(* IEC 61131-3 sources: STAR-PLC-Agent/results/raw/four_group_20261114/star_terra/PUB008/generation/sim_00, 1 file *)

(* ---- test_program.st ---- *)
PROGRAM PLC_PRG
VAR
 BenchStep : UDINT := 0;
 BenchCalls : UDINT := 0;
 BenchDone : BOOL := FALSE;
 BenchUut0 : FB_Task;
 BenchUut1 : FB_Task;
 Binding_0_analogValues : ARRAY[1..14] OF INT;
 Binding_0_channels : ARRAY[1..14] OF ST_AnalogChannel;
 Binding_1_analogValues : ARRAY[1..10] OF INT;
 Binding_1_channels : ARRAY[1..9] OF ST_AnalogChannel;
 TraceIn_count : ARRAY[0..3] OF DINT;
 TraceOut_analogValues_1 : ARRAY[0..3] OF INT;
 TraceOut_analogValues_2 : ARRAY[0..3] OF INT;
 TraceOut_analogValues_3 : ARRAY[0..3] OF INT;
 TraceOut_analogValues_4 : ARRAY[0..3] OF INT;
 TraceOut_analogValues_5 : ARRAY[0..3] OF INT;
 TraceOut_analogValues_6 : ARRAY[0..3] OF INT;
 TraceOut_analogValues_7 : ARRAY[0..3] OF INT;
 TraceOut_analogValues_8 : ARRAY[0..3] OF INT;
 TraceOut_analogValues_9 : ARRAY[0..3] OF INT;
 TraceOut_analogValues_10 : ARRAY[0..3] OF INT;
 TraceOut_analogValues_11 : ARRAY[0..3] OF INT;
 TraceOut_analogValues_12 : ARRAY[0..3] OF INT;
 TraceOut_analogValues_13 : ARRAY[0..3] OF INT;
 TraceOut_analogValues_14 : ARRAY[0..3] OF INT;
 TraceOut_channels_1_enable : ARRAY[0..3] OF BOOL;
 TraceOut_channels_1_hiLIM : ARRAY[0..3] OF REAL;
 TraceOut_channels_1_loLIM : ARRAY[0..3] OF REAL;
 TraceOut_channels_1_bipolar : ARRAY[0..3] OF BOOL;
 TraceOut_channels_1_measuringMode : ARRAY[0..3] OF INT;
 TraceOut_channels_1_retVal : ARRAY[0..3] OF WORD;
 TraceOut_channels_1_outputValue : ARRAY[0..3] OF REAL;
 TraceOut_channels_2_enable : ARRAY[0..3] OF BOOL;
 TraceOut_channels_2_hiLIM : ARRAY[0..3] OF REAL;
 TraceOut_channels_2_loLIM : ARRAY[0..3] OF REAL;
 TraceOut_channels_2_bipolar : ARRAY[0..3] OF BOOL;
 TraceOut_channels_2_measuringMode : ARRAY[0..3] OF INT;
 TraceOut_channels_2_retVal : ARRAY[0..3] OF WORD;
 TraceOut_channels_2_outputValue : ARRAY[0..3] OF REAL;
 TraceOut_channels_3_enable : ARRAY[0..3] OF BOOL;
 TraceOut_channels_3_hiLIM : ARRAY[0..3] OF REAL;
 TraceOut_channels_3_loLIM : ARRAY[0..3] OF REAL;
 TraceOut_channels_3_bipolar : ARRAY[0..3] OF BOOL;
 TraceOut_channels_3_measuringMode : ARRAY[0..3] OF INT;
 TraceOut_channels_3_retVal : ARRAY[0..3] OF WORD;
 TraceOut_channels_3_outputValue : ARRAY[0..3] OF REAL;
 TraceOut_channels_4_enable : ARRAY[0..3] OF BOOL;
 TraceOut_channels_4_hiLIM : ARRAY[0..3] OF REAL;
 TraceOut_channels_4_loLIM : ARRAY[0..3] OF REAL;
 TraceOut_channels_4_bipolar : ARRAY[0..3] OF BOOL;
 TraceOut_channels_4_measuringMode : ARRAY[0..3] OF INT;
 TraceOut_channels_4_retVal : ARRAY[0..3] OF WORD;
 TraceOut_channels_4_outputValue : ARRAY[0..3] OF REAL;
 TraceOut_channels_5_enable : ARRAY[0..3] OF BOOL;
 TraceOut_channels_5_hiLIM : ARRAY[0..3] OF REAL;
 TraceOut_channels_5_loLIM : ARRAY[0..3] OF REAL;
 TraceOut_channels_5_bipolar : ARRAY[0..3] OF BOOL;
 TraceOut_channels_5_measuringMode : ARRAY[0..3] OF INT;
 TraceOut_channels_5_retVal : ARRAY[0..3] OF WORD;
 TraceOut_channels_5_outputValue : ARRAY[0..3] OF REAL;
 TraceOut_channels_6_enable : ARRAY[0..3] OF BOOL;
 TraceOut_channels_6_hiLIM : ARRAY[0..3] OF REAL;
 TraceOut_channels_6_loLIM : ARRAY[0..3] OF REAL;
 TraceOut_channels_6_bipolar : ARRAY[0..3] OF BOOL;
 TraceOut_channels_6_measuringMode : ARRAY[0..3] OF INT;
 TraceOut_channels_6_retVal : ARRAY[0..3] OF WORD;
 TraceOut_channels_6_outputValue : ARRAY[0..3] OF REAL;
 TraceOut_channels_7_enable : ARRAY[0..3] OF BOOL;
 TraceOut_channels_7_hiLIM : ARRAY[0..3] OF REAL;
 TraceOut_channels_7_loLIM : ARRAY[0..3] OF REAL;
 TraceOut_channels_7_bipolar : ARRAY[0..3] OF BOOL;
 TraceOut_channels_7_measuringMode : ARRAY[0..3] OF INT;
 TraceOut_channels_7_retVal : ARRAY[0..3] OF WORD;
 TraceOut_channels_7_outputValue : ARRAY[0..3] OF REAL;
 TraceOut_channels_8_enable : ARRAY[0..3] OF BOOL;
 TraceOut_channels_8_hiLIM : ARRAY[0..3] OF REAL;
 TraceOut_channels_8_loLIM : ARRAY[0..3] OF REAL;
 TraceOut_channels_8_bipolar : ARRAY[0..3] OF BOOL;
 TraceOut_channels_8_measuringMode : ARRAY[0..3] OF INT;
 TraceOut_channels_8_retVal : ARRAY[0..3] OF WORD;
 TraceOut_channels_8_outputValue : ARRAY[0..3] OF REAL;
 TraceOut_channels_9_enable : ARRAY[0..3] OF BOOL;
 TraceOut_channels_9_hiLIM : ARRAY[0..3] OF REAL;
 TraceOut_channels_9_loLIM : ARRAY[0..3] OF REAL;
 TraceOut_channels_9_bipolar : ARRAY[0..3] OF BOOL;
 TraceOut_channels_9_measuringMode : ARRAY[0..3] OF INT;
 TraceOut_channels_9_retVal : ARRAY[0..3] OF WORD;
 TraceOut_channels_9_outputValue : ARRAY[0..3] OF REAL;
 TraceOut_channels_10_enable : ARRAY[0..3] OF BOOL;
 TraceOut_channels_10_hiLIM : ARRAY[0..3] OF REAL;
 TraceOut_channels_10_loLIM : ARRAY[0..3] OF REAL;
 TraceOut_channels_10_bipolar : ARRAY[0..3] OF BOOL;
 TraceOut_channels_10_measuringMode : ARRAY[0..3] OF INT;
 TraceOut_channels_10_retVal : ARRAY[0..3] OF WORD;
 TraceOut_channels_10_outputValue : ARRAY[0..3] OF REAL;
 TraceOut_channels_11_enable : ARRAY[0..3] OF BOOL;
 TraceOut_channels_11_hiLIM : ARRAY[0..3] OF REAL;
 TraceOut_channels_11_loLIM : ARRAY[0..3] OF REAL;
 TraceOut_channels_11_bipolar : ARRAY[0..3] OF BOOL;
 TraceOut_channels_11_measuringMode : ARRAY[0..3] OF INT;
 TraceOut_channels_11_retVal : ARRAY[0..3] OF WORD;
 TraceOut_channels_11_outputValue : ARRAY[0..3] OF REAL;
 TraceOut_channels_12_enable : ARRAY[0..3] OF BOOL;
 TraceOut_channels_12_hiLIM : ARRAY[0..3] OF REAL;
 TraceOut_channels_12_loLIM : ARRAY[0..3] OF REAL;
 TraceOut_channels_12_bipolar : ARRAY[0..3] OF BOOL;
 TraceOut_channels_12_measuringMode : ARRAY[0..3] OF INT;
 TraceOut_channels_12_retVal : ARRAY[0..3] OF WORD;
 TraceOut_channels_12_outputValue : ARRAY[0..3] OF REAL;
 TraceOut_channels_13_enable : ARRAY[0..3] OF BOOL;
 TraceOut_channels_13_hiLIM : ARRAY[0..3] OF REAL;
 TraceOut_channels_13_loLIM : ARRAY[0..3] OF REAL;
 TraceOut_channels_13_bipolar : ARRAY[0..3] OF BOOL;
 TraceOut_channels_13_measuringMode : ARRAY[0..3] OF INT;
 TraceOut_channels_13_retVal : ARRAY[0..3] OF WORD;
 TraceOut_channels_13_outputValue : ARRAY[0..3] OF REAL;
 TraceOut_channels_14_enable : ARRAY[0..3] OF BOOL;
 TraceOut_channels_14_hiLIM : ARRAY[0..3] OF REAL;
 TraceOut_channels_14_loLIM : ARRAY[0..3] OF REAL;
 TraceOut_channels_14_bipolar : ARRAY[0..3] OF BOOL;
 TraceOut_channels_14_measuringMode : ARRAY[0..3] OF INT;
 TraceOut_channels_14_retVal : ARRAY[0..3] OF WORD;
 TraceOut_channels_14_outputValue : ARRAY[0..3] OF REAL;
 TraceInIO_analogValues_e0_INT : ARRAY[0..3] OF INT;
 TraceInIO_analogValues_e1_INT : ARRAY[0..3] OF INT;
 TraceInIO_analogValues_e2_INT : ARRAY[0..3] OF INT;
 TraceInIO_analogValues_e3_INT : ARRAY[0..3] OF INT;
 TraceInIO_analogValues_e4_INT : ARRAY[0..3] OF INT;
 TraceInIO_analogValues_e5_INT : ARRAY[0..3] OF INT;
 TraceInIO_analogValues_e6_INT : ARRAY[0..3] OF INT;
 TraceInIO_analogValues_e7_INT : ARRAY[0..3] OF INT;
 TraceInIO_analogValues_e8_INT : ARRAY[0..3] OF INT;
 TraceInIO_analogValues_e9_INT : ARRAY[0..3] OF INT;
 TraceInIO_analogValues_e10_INT : ARRAY[0..3] OF INT;
 TraceInIO_analogValues_e11_INT : ARRAY[0..3] OF INT;
 TraceInIO_analogValues_e12_INT : ARRAY[0..3] OF INT;
 TraceInIO_analogValues_e13_INT : ARRAY[0..3] OF INT;
 TraceInIO_channels_e0_enable_BOOL : ARRAY[0..3] OF BOOL;
 TraceInIO_channels_e0_hiLIM_REAL : ARRAY[0..3] OF REAL;
 TraceInIO_channels_e0_loLIM_REAL : ARRAY[0..3] OF REAL;
 TraceInIO_channels_e0_bipolar_BOOL : ARRAY[0..3] OF BOOL;
 TraceInIO_channels_e0_measuringMode_INT : ARRAY[0..3] OF INT;
 TraceInIO_channels_e0_retVal_WORD : ARRAY[0..3] OF WORD;
 TraceInIO_channels_e0_outputValue_REAL : ARRAY[0..3] OF REAL;
 TraceInIO_channels_e1_enable_BOOL : ARRAY[0..3] OF BOOL;
 TraceInIO_channels_e1_hiLIM_REAL : ARRAY[0..3] OF REAL;
 TraceInIO_channels_e1_loLIM_REAL : ARRAY[0..3] OF REAL;
 TraceInIO_channels_e1_bipolar_BOOL : ARRAY[0..3] OF BOOL;
 TraceInIO_channels_e1_measuringMode_INT : ARRAY[0..3] OF INT;
 TraceInIO_channels_e1_retVal_WORD : ARRAY[0..3] OF WORD;
 TraceInIO_channels_e1_outputValue_REAL : ARRAY[0..3] OF REAL;
 TraceInIO_channels_e2_enable_BOOL : ARRAY[0..3] OF BOOL;
 TraceInIO_channels_e2_hiLIM_REAL : ARRAY[0..3] OF REAL;
 TraceInIO_channels_e2_loLIM_REAL : ARRAY[0..3] OF REAL;
 TraceInIO_channels_e2_bipolar_BOOL : ARRAY[0..3] OF BOOL;
 TraceInIO_channels_e2_measuringMode_INT : ARRAY[0..3] OF INT;
 TraceInIO_channels_e2_retVal_WORD : ARRAY[0..3] OF WORD;
 TraceInIO_channels_e2_outputValue_REAL : ARRAY[0..3] OF REAL;
 TraceInIO_channels_e3_enable_BOOL : ARRAY[0..3] OF BOOL;
 TraceInIO_channels_e3_hiLIM_REAL : ARRAY[0..3] OF REAL;
 TraceInIO_channels_e3_loLIM_REAL : ARRAY[0..3] OF REAL;
 TraceInIO_channels_e3_bipolar_BOOL : ARRAY[0..3] OF BOOL;
 TraceInIO_channels_e3_measuringMode_INT : ARRAY[0..3] OF INT;
 TraceInIO_channels_e3_retVal_WORD : ARRAY[0..3] OF WORD;
 TraceInIO_channels_e3_outputValue_REAL : ARRAY[0..3] OF REAL;
 TraceInIO_channels_e4_enable_BOOL : ARRAY[0..3] OF BOOL;
 TraceInIO_channels_e4_hiLIM_REAL : ARRAY[0..3] OF REAL;
 TraceInIO_channels_e4_loLIM_REAL : ARRAY[0..3] OF REAL;
 TraceInIO_channels_e4_bipolar_BOOL : ARRAY[0..3] OF BOOL;
 TraceInIO_channels_e4_measuringMode_INT : ARRAY[0..3] OF INT;
 TraceInIO_channels_e4_retVal_WORD : ARRAY[0..3] OF WORD;
 TraceInIO_channels_e4_outputValue_REAL : ARRAY[0..3] OF REAL;
 TraceInIO_channels_e5_enable_BOOL : ARRAY[0..3] OF BOOL;
 TraceInIO_channels_e5_hiLIM_REAL : ARRAY[0..3] OF REAL;
 TraceInIO_channels_e5_loLIM_REAL : ARRAY[0..3] OF REAL;
 TraceInIO_channels_e5_bipolar_BOOL : ARRAY[0..3] OF BOOL;
 TraceInIO_channels_e5_measuringMode_INT : ARRAY[0..3] OF INT;
 TraceInIO_channels_e5_retVal_WORD : ARRAY[0..3] OF WORD;
 TraceInIO_channels_e5_outputValue_REAL : ARRAY[0..3] OF REAL;
 TraceInIO_channels_e6_enable_BOOL : ARRAY[0..3] OF BOOL;
 TraceInIO_channels_e6_hiLIM_REAL : ARRAY[0..3] OF REAL;
 TraceInIO_channels_e6_loLIM_REAL : ARRAY[0..3] OF REAL;
 TraceInIO_channels_e6_bipolar_BOOL : ARRAY[0..3] OF BOOL;
 TraceInIO_channels_e6_measuringMode_INT : ARRAY[0..3] OF INT;
 TraceInIO_channels_e6_retVal_WORD : ARRAY[0..3] OF WORD;
 TraceInIO_channels_e6_outputValue_REAL : ARRAY[0..3] OF REAL;
 TraceInIO_channels_e7_enable_BOOL : ARRAY[0..3] OF BOOL;
 TraceInIO_channels_e7_hiLIM_REAL : ARRAY[0..3] OF REAL;
 TraceInIO_channels_e7_loLIM_REAL : ARRAY[0..3] OF REAL;
 TraceInIO_channels_e7_bipolar_BOOL : ARRAY[0..3] OF BOOL;
 TraceInIO_channels_e7_measuringMode_INT : ARRAY[0..3] OF INT;
 TraceInIO_channels_e7_retVal_WORD : ARRAY[0..3] OF WORD;
 TraceInIO_channels_e7_outputValue_REAL : ARRAY[0..3] OF REAL;
 TraceInIO_channels_e8_enable_BOOL : ARRAY[0..3] OF BOOL;
 TraceInIO_channels_e8_hiLIM_REAL : ARRAY[0..3] OF REAL;
 TraceInIO_channels_e8_loLIM_REAL : ARRAY[0..3] OF REAL;
 TraceInIO_channels_e8_bipolar_BOOL : ARRAY[0..3] OF BOOL;
 TraceInIO_channels_e8_measuringMode_INT : ARRAY[0..3] OF INT;
 TraceInIO_channels_e8_retVal_WORD : ARRAY[0..3] OF WORD;
 TraceInIO_channels_e8_outputValue_REAL : ARRAY[0..3] OF REAL;
 TraceInIO_channels_e9_enable_BOOL : ARRAY[0..3] OF BOOL;
 TraceInIO_channels_e9_hiLIM_REAL : ARRAY[0..3] OF REAL;
 TraceInIO_channels_e9_loLIM_REAL : ARRAY[0..3] OF REAL;
 TraceInIO_channels_e9_bipolar_BOOL : ARRAY[0..3] OF BOOL;
 TraceInIO_channels_e9_measuringMode_INT : ARRAY[0..3] OF INT;
 TraceInIO_channels_e9_retVal_WORD : ARRAY[0..3] OF WORD;
 TraceInIO_channels_e9_outputValue_REAL : ARRAY[0..3] OF REAL;
 TraceInIO_channels_e10_enable_BOOL : ARRAY[0..3] OF BOOL;
 TraceInIO_channels_e10_hiLIM_REAL : ARRAY[0..3] OF REAL;
 TraceInIO_channels_e10_loLIM_REAL : ARRAY[0..3] OF REAL;
 TraceInIO_channels_e10_bipolar_BOOL : ARRAY[0..3] OF BOOL;
 TraceInIO_channels_e10_measuringMode_INT : ARRAY[0..3] OF INT;
 TraceInIO_channels_e10_retVal_WORD : ARRAY[0..3] OF WORD;
 TraceInIO_channels_e10_outputValue_REAL : ARRAY[0..3] OF REAL;
 TraceInIO_channels_e11_enable_BOOL : ARRAY[0..3] OF BOOL;
 TraceInIO_channels_e11_hiLIM_REAL : ARRAY[0..3] OF REAL;
 TraceInIO_channels_e11_loLIM_REAL : ARRAY[0..3] OF REAL;
 TraceInIO_channels_e11_bipolar_BOOL : ARRAY[0..3] OF BOOL;
 TraceInIO_channels_e11_measuringMode_INT : ARRAY[0..3] OF INT;
 TraceInIO_channels_e11_retVal_WORD : ARRAY[0..3] OF WORD;
 TraceInIO_channels_e11_outputValue_REAL : ARRAY[0..3] OF REAL;
 TraceInIO_channels_e12_enable_BOOL : ARRAY[0..3] OF BOOL;
 TraceInIO_channels_e12_hiLIM_REAL : ARRAY[0..3] OF REAL;
 TraceInIO_channels_e12_loLIM_REAL : ARRAY[0..3] OF REAL;
 TraceInIO_channels_e12_bipolar_BOOL : ARRAY[0..3] OF BOOL;
 TraceInIO_channels_e12_measuringMode_INT : ARRAY[0..3] OF INT;
 TraceInIO_channels_e12_retVal_WORD : ARRAY[0..3] OF WORD;
 TraceInIO_channels_e12_outputValue_REAL : ARRAY[0..3] OF REAL;
 TraceInIO_channels_e13_enable_BOOL : ARRAY[0..3] OF BOOL;
 TraceInIO_channels_e13_hiLIM_REAL : ARRAY[0..3] OF REAL;
 TraceInIO_channels_e13_loLIM_REAL : ARRAY[0..3] OF REAL;
 TraceInIO_channels_e13_bipolar_BOOL : ARRAY[0..3] OF BOOL;
 TraceInIO_channels_e13_measuringMode_INT : ARRAY[0..3] OF INT;
 TraceInIO_channels_e13_retVal_WORD : ARRAY[0..3] OF WORD;
 TraceInIO_channels_e13_outputValue_REAL : ARRAY[0..3] OF REAL;
END_VAR

IF NOT BenchDone THEN
 CASE BenchStep OF
 0:
   Binding_0_analogValues[1] := INT#0;
   Binding_0_analogValues[2] := INT#27648;
   Binding_0_analogValues[3] := INT#13824;
   Binding_0_analogValues[4] := INT#-27648;
   Binding_0_analogValues[5] := INT#-27648;
   Binding_0_analogValues[6] := INT#0;
   Binding_0_analogValues[7] := INT#27648;
   Binding_0_analogValues[8] := INT#13824;
   Binding_0_analogValues[9] := INT#1234;
   Binding_0_analogValues[10] := INT#-2345;
   Binding_0_analogValues[11] := INT#123;
   Binding_0_analogValues[12] := INT#-1;
   Binding_0_analogValues[13] := INT#333;
   Binding_0_analogValues[14] := INT#222;
   Binding_0_channels[1].enable := TRUE;
   Binding_0_channels[1].hiLIM := REAL#110.0;
   Binding_0_channels[1].loLIM := REAL#10.0;
   Binding_0_channels[1].bipolar := FALSE;
   Binding_0_channels[1].measuringMode := INT#0;
   Binding_0_channels[1].retVal := WORD#11;
   Binding_0_channels[1].outputValue := REAL#-1.0;
   Binding_0_channels[2].enable := TRUE;
   Binding_0_channels[2].hiLIM := REAL#110.0;
   Binding_0_channels[2].loLIM := REAL#10.0;
   Binding_0_channels[2].bipolar := FALSE;
   Binding_0_channels[2].measuringMode := INT#0;
   Binding_0_channels[2].retVal := WORD#12;
   Binding_0_channels[2].outputValue := REAL#-2.0;
   Binding_0_channels[3].enable := TRUE;
   Binding_0_channels[3].hiLIM := REAL#110.0;
   Binding_0_channels[3].loLIM := REAL#10.0;
   Binding_0_channels[3].bipolar := FALSE;
   Binding_0_channels[3].measuringMode := INT#0;
   Binding_0_channels[3].retVal := WORD#13;
   Binding_0_channels[3].outputValue := REAL#-3.0;
   Binding_0_channels[4].enable := TRUE;
   Binding_0_channels[4].hiLIM := REAL#110.0;
   Binding_0_channels[4].loLIM := REAL#10.0;
   Binding_0_channels[4].bipolar := FALSE;
   Binding_0_channels[4].measuringMode := INT#0;
   Binding_0_channels[4].retVal := WORD#14;
   Binding_0_channels[4].outputValue := REAL#-4.0;
   Binding_0_channels[5].enable := TRUE;
   Binding_0_channels[5].hiLIM := REAL#30.0;
   Binding_0_channels[5].loLIM := REAL#-20.0;
   Binding_0_channels[5].bipolar := TRUE;
   Binding_0_channels[5].measuringMode := INT#0;
   Binding_0_channels[5].retVal := WORD#15;
   Binding_0_channels[5].outputValue := REAL#-5.0;
   Binding_0_channels[6].enable := TRUE;
   Binding_0_channels[6].hiLIM := REAL#30.0;
   Binding_0_channels[6].loLIM := REAL#-20.0;
   Binding_0_channels[6].bipolar := TRUE;
   Binding_0_channels[6].measuringMode := INT#0;
   Binding_0_channels[6].retVal := WORD#16;
   Binding_0_channels[6].outputValue := REAL#-6.0;
   Binding_0_channels[7].enable := TRUE;
   Binding_0_channels[7].hiLIM := REAL#30.0;
   Binding_0_channels[7].loLIM := REAL#-20.0;
   Binding_0_channels[7].bipolar := TRUE;
   Binding_0_channels[7].measuringMode := INT#0;
   Binding_0_channels[7].retVal := WORD#17;
   Binding_0_channels[7].outputValue := REAL#-7.0;
   Binding_0_channels[8].enable := TRUE;
   Binding_0_channels[8].hiLIM := REAL#30.0;
   Binding_0_channels[8].loLIM := REAL#-20.0;
   Binding_0_channels[8].bipolar := TRUE;
   Binding_0_channels[8].measuringMode := INT#0;
   Binding_0_channels[8].retVal := WORD#18;
   Binding_0_channels[8].outputValue := REAL#-8.0;
   Binding_0_channels[9].enable := TRUE;
   Binding_0_channels[9].hiLIM := REAL#1.0;
   Binding_0_channels[9].loLIM := REAL#0.0;
   Binding_0_channels[9].bipolar := FALSE;
   Binding_0_channels[9].measuringMode := INT#1;
   Binding_0_channels[9].retVal := WORD#19;
   Binding_0_channels[9].outputValue := REAL#-9.0;
   Binding_0_channels[10].enable := TRUE;
   Binding_0_channels[10].hiLIM := REAL#1.0;
   Binding_0_channels[10].loLIM := REAL#0.0;
   Binding_0_channels[10].bipolar := TRUE;
   Binding_0_channels[10].measuringMode := INT#1;
   Binding_0_channels[10].retVal := WORD#20;
   Binding_0_channels[10].outputValue := REAL#-10.0;
   Binding_0_channels[11].enable := TRUE;
   Binding_0_channels[11].hiLIM := REAL#1.0;
   Binding_0_channels[11].loLIM := REAL#0.0;
   Binding_0_channels[11].bipolar := FALSE;
   Binding_0_channels[11].measuringMode := INT#2;
   Binding_0_channels[11].retVal := WORD#21;
   Binding_0_channels[11].outputValue := REAL#-11.0;
   Binding_0_channels[12].enable := TRUE;
   Binding_0_channels[12].hiLIM := REAL#1.0;
   Binding_0_channels[12].loLIM := REAL#0.0;
   Binding_0_channels[12].bipolar := TRUE;
   Binding_0_channels[12].measuringMode := INT#2;
   Binding_0_channels[12].retVal := WORD#22;
   Binding_0_channels[12].outputValue := REAL#-12.0;
   Binding_0_channels[13].enable := FALSE;
   Binding_0_channels[13].hiLIM := REAL#0.0;
   Binding_0_channels[13].loLIM := REAL#0.0;
   Binding_0_channels[13].bipolar := TRUE;
   Binding_0_channels[13].measuringMode := INT#99;
   Binding_0_channels[13].retVal := WORD#23;
   Binding_0_channels[13].outputValue := REAL#-13.0;
   Binding_0_channels[14].enable := TRUE;
   Binding_0_channels[14].hiLIM := REAL#100.0;
   Binding_0_channels[14].loLIM := REAL#0.0;
   Binding_0_channels[14].bipolar := FALSE;
   Binding_0_channels[14].measuringMode := INT#0;
   Binding_0_channels[14].retVal := WORD#24;
   Binding_0_channels[14].outputValue := REAL#-14.0;
   BenchUut0.count := DINT#13;
   TraceIn_count[0] := BenchUut0.count;
   TraceInIO_analogValues_e0_INT[0] := Binding_0_analogValues[1];
   TraceInIO_analogValues_e1_INT[0] := Binding_0_analogValues[2];
   TraceInIO_analogValues_e2_INT[0] := Binding_0_analogValues[3];
   TraceInIO_analogValues_e3_INT[0] := Binding_0_analogValues[4];
   TraceInIO_analogValues_e4_INT[0] := Binding_0_analogValues[5];
   TraceInIO_analogValues_e5_INT[0] := Binding_0_analogValues[6];
   TraceInIO_analogValues_e6_INT[0] := Binding_0_analogValues[7];
   TraceInIO_analogValues_e7_INT[0] := Binding_0_analogValues[8];
   TraceInIO_analogValues_e8_INT[0] := Binding_0_analogValues[9];
   TraceInIO_analogValues_e9_INT[0] := Binding_0_analogValues[10];
   TraceInIO_analogValues_e10_INT[0] := Binding_0_analogValues[11];
   TraceInIO_analogValues_e11_INT[0] := Binding_0_analogValues[12];
   TraceInIO_analogValues_e12_INT[0] := Binding_0_analogValues[13];
   TraceInIO_analogValues_e13_INT[0] := Binding_0_analogValues[14];
   TraceInIO_channels_e0_enable_BOOL[0] := Binding_0_channels[1].enable;
   TraceInIO_channels_e0_hiLIM_REAL[0] := Binding_0_channels[1].hiLIM;
   TraceInIO_channels_e0_loLIM_REAL[0] := Binding_0_channels[1].loLIM;
   TraceInIO_channels_e0_bipolar_BOOL[0] := Binding_0_channels[1].bipolar;
   TraceInIO_channels_e0_measuringMode_INT[0] := Binding_0_channels[1].measuringMode;
   TraceInIO_channels_e0_retVal_WORD[0] := Binding_0_channels[1].retVal;
   TraceInIO_channels_e0_outputValue_REAL[0] := Binding_0_channels[1].outputValue;
   TraceInIO_channels_e1_enable_BOOL[0] := Binding_0_channels[2].enable;
   TraceInIO_channels_e1_hiLIM_REAL[0] := Binding_0_channels[2].hiLIM;
   TraceInIO_channels_e1_loLIM_REAL[0] := Binding_0_channels[2].loLIM;
   TraceInIO_channels_e1_bipolar_BOOL[0] := Binding_0_channels[2].bipolar;
   TraceInIO_channels_e1_measuringMode_INT[0] := Binding_0_channels[2].measuringMode;
   TraceInIO_channels_e1_retVal_WORD[0] := Binding_0_channels[2].retVal;
   TraceInIO_channels_e1_outputValue_REAL[0] := Binding_0_channels[2].outputValue;
   TraceInIO_channels_e2_enable_BOOL[0] := Binding_0_channels[3].enable;
   TraceInIO_channels_e2_hiLIM_REAL[0] := Binding_0_channels[3].hiLIM;
   TraceInIO_channels_e2_loLIM_REAL[0] := Binding_0_channels[3].loLIM;
   TraceInIO_channels_e2_bipolar_BOOL[0] := Binding_0_channels[3].bipolar;
   TraceInIO_channels_e2_measuringMode_INT[0] := Binding_0_channels[3].measuringMode;
   TraceInIO_channels_e2_retVal_WORD[0] := Binding_0_channels[3].retVal;
   TraceInIO_channels_e2_outputValue_REAL[0] := Binding_0_channels[3].outputValue;
   TraceInIO_channels_e3_enable_BOOL[0] := Binding_0_channels[4].enable;
   TraceInIO_channels_e3_hiLIM_REAL[0] := Binding_0_channels[4].hiLIM;
   TraceInIO_channels_e3_loLIM_REAL[0] := Binding_0_channels[4].loLIM;
   TraceInIO_channels_e3_bipolar_BOOL[0] := Binding_0_channels[4].bipolar;
   TraceInIO_channels_e3_measuringMode_INT[0] := Binding_0_channels[4].measuringMode;
   TraceInIO_channels_e3_retVal_WORD[0] := Binding_0_channels[4].retVal;
   TraceInIO_channels_e3_outputValue_REAL[0] := Binding_0_channels[4].outputValue;
   TraceInIO_channels_e4_enable_BOOL[0] := Binding_0_channels[5].enable;
   TraceInIO_channels_e4_hiLIM_REAL[0] := Binding_0_channels[5].hiLIM;
   TraceInIO_channels_e4_loLIM_REAL[0] := Binding_0_channels[5].loLIM;
   TraceInIO_channels_e4_bipolar_BOOL[0] := Binding_0_channels[5].bipolar;
   TraceInIO_channels_e4_measuringMode_INT[0] := Binding_0_channels[5].measuringMode;
   TraceInIO_channels_e4_retVal_WORD[0] := Binding_0_channels[5].retVal;
   TraceInIO_channels_e4_outputValue_REAL[0] := Binding_0_channels[5].outputValue;
   TraceInIO_channels_e5_enable_BOOL[0] := Binding_0_channels[6].enable;
   TraceInIO_channels_e5_hiLIM_REAL[0] := Binding_0_channels[6].hiLIM;
   TraceInIO_channels_e5_loLIM_REAL[0] := Binding_0_channels[6].loLIM;
   TraceInIO_channels_e5_bipolar_BOOL[0] := Binding_0_channels[6].bipolar;
   TraceInIO_channels_e5_measuringMode_INT[0] := Binding_0_channels[6].measuringMode;
   TraceInIO_channels_e5_retVal_WORD[0] := Binding_0_channels[6].retVal;
   TraceInIO_channels_e5_outputValue_REAL[0] := Binding_0_channels[6].outputValue;
   TraceInIO_channels_e6_enable_BOOL[0] := Binding_0_channels[7].enable;
   TraceInIO_channels_e6_hiLIM_REAL[0] := Binding_0_channels[7].hiLIM;
   TraceInIO_channels_e6_loLIM_REAL[0] := Binding_0_channels[7].loLIM;
   TraceInIO_channels_e6_bipolar_BOOL[0] := Binding_0_channels[7].bipolar;
   TraceInIO_channels_e6_measuringMode_INT[0] := Binding_0_channels[7].measuringMode;
   TraceInIO_channels_e6_retVal_WORD[0] := Binding_0_channels[7].retVal;
   TraceInIO_channels_e6_outputValue_REAL[0] := Binding_0_channels[7].outputValue;
   TraceInIO_channels_e7_enable_BOOL[0] := Binding_0_channels[8].enable;
   TraceInIO_channels_e7_hiLIM_REAL[0] := Binding_0_channels[8].hiLIM;
   TraceInIO_channels_e7_loLIM_REAL[0] := Binding_0_channels[8].loLIM;
   TraceInIO_channels_e7_bipolar_BOOL[0] := Binding_0_channels[8].bipolar;
   TraceInIO_channels_e7_measuringMode_INT[0] := Binding_0_channels[8].measuringMode;
   TraceInIO_channels_e7_retVal_WORD[0] := Binding_0_channels[8].retVal;
   TraceInIO_channels_e7_outputValue_REAL[0] := Binding_0_channels[8].outputValue;
   TraceInIO_channels_e8_enable_BOOL[0] := Binding_0_channels[9].enable;
   TraceInIO_channels_e8_hiLIM_REAL[0] := Binding_0_channels[9].hiLIM;
   TraceInIO_channels_e8_loLIM_REAL[0] := Binding_0_channels[9].loLIM;
   TraceInIO_channels_e8_bipolar_BOOL[0] := Binding_0_channels[9].bipolar;
   TraceInIO_channels_e8_measuringMode_INT[0] := Binding_0_channels[9].measuringMode;
   TraceInIO_channels_e8_retVal_WORD[0] := Binding_0_channels[9].retVal;
   TraceInIO_channels_e8_outputValue_REAL[0] := Binding_0_channels[9].outputValue;
   TraceInIO_channels_e9_enable_BOOL[0] := Binding_0_channels[10].enable;
   TraceInIO_channels_e9_hiLIM_REAL[0] := Binding_0_channels[10].hiLIM;
   TraceInIO_channels_e9_loLIM_REAL[0] := Binding_0_channels[10].loLIM;
   TraceInIO_channels_e9_bipolar_BOOL[0] := Binding_0_channels[10].bipolar;
   TraceInIO_channels_e9_measuringMode_INT[0] := Binding_0_channels[10].measuringMode;
   TraceInIO_channels_e9_retVal_WORD[0] := Binding_0_channels[10].retVal;
   TraceInIO_channels_e9_outputValue_REAL[0] := Binding_0_channels[10].outputValue;
   TraceInIO_channels_e10_enable_BOOL[0] := Binding_0_channels[11].enable;
   TraceInIO_channels_e10_hiLIM_REAL[0] := Binding_0_channels[11].hiLIM;
   TraceInIO_channels_e10_loLIM_REAL[0] := Binding_0_channels[11].loLIM;
   TraceInIO_channels_e10_bipolar_BOOL[0] := Binding_0_channels[11].bipolar;
   TraceInIO_channels_e10_measuringMode_INT[0] := Binding_0_channels[11].measuringMode;
   TraceInIO_channels_e10_retVal_WORD[0] := Binding_0_channels[11].retVal;
   TraceInIO_channels_e10_outputValue_REAL[0] := Binding_0_channels[11].outputValue;
   TraceInIO_channels_e11_enable_BOOL[0] := Binding_0_channels[12].enable;
   TraceInIO_channels_e11_hiLIM_REAL[0] := Binding_0_channels[12].hiLIM;
   TraceInIO_channels_e11_loLIM_REAL[0] := Binding_0_channels[12].loLIM;
   TraceInIO_channels_e11_bipolar_BOOL[0] := Binding_0_channels[12].bipolar;
   TraceInIO_channels_e11_measuringMode_INT[0] := Binding_0_channels[12].measuringMode;
   TraceInIO_channels_e11_retVal_WORD[0] := Binding_0_channels[12].retVal;
   TraceInIO_channels_e11_outputValue_REAL[0] := Binding_0_channels[12].outputValue;
   TraceInIO_channels_e12_enable_BOOL[0] := Binding_0_channels[13].enable;
   TraceInIO_channels_e12_hiLIM_REAL[0] := Binding_0_channels[13].hiLIM;
   TraceInIO_channels_e12_loLIM_REAL[0] := Binding_0_channels[13].loLIM;
   TraceInIO_channels_e12_bipolar_BOOL[0] := Binding_0_channels[13].bipolar;
   TraceInIO_channels_e12_measuringMode_INT[0] := Binding_0_channels[13].measuringMode;
   TraceInIO_channels_e12_retVal_WORD[0] := Binding_0_channels[13].retVal;
   TraceInIO_channels_e12_outputValue_REAL[0] := Binding_0_channels[13].outputValue;
   TraceInIO_channels_e13_enable_BOOL[0] := Binding_0_channels[14].enable;
   TraceInIO_channels_e13_hiLIM_REAL[0] := Binding_0_channels[14].hiLIM;
   TraceInIO_channels_e13_loLIM_REAL[0] := Binding_0_channels[14].loLIM;
   TraceInIO_channels_e13_bipolar_BOOL[0] := Binding_0_channels[14].bipolar;
   TraceInIO_channels_e13_measuringMode_INT[0] := Binding_0_channels[14].measuringMode;
   TraceInIO_channels_e13_retVal_WORD[0] := Binding_0_channels[14].retVal;
   TraceInIO_channels_e13_outputValue_REAL[0] := Binding_0_channels[14].outputValue;
   BenchUut0(analogValues := Binding_0_analogValues, channels := Binding_0_channels);
   TraceOut_analogValues_1[0] := Binding_0_analogValues[1];
   TraceOut_analogValues_2[0] := Binding_0_analogValues[2];
   TraceOut_analogValues_3[0] := Binding_0_analogValues[3];
   TraceOut_analogValues_4[0] := Binding_0_analogValues[4];
   TraceOut_analogValues_5[0] := Binding_0_analogValues[5];
   TraceOut_analogValues_6[0] := Binding_0_analogValues[6];
   TraceOut_analogValues_7[0] := Binding_0_analogValues[7];
   TraceOut_analogValues_8[0] := Binding_0_analogValues[8];
   TraceOut_analogValues_9[0] := Binding_0_analogValues[9];
   TraceOut_analogValues_10[0] := Binding_0_analogValues[10];
   TraceOut_analogValues_11[0] := Binding_0_analogValues[11];
   TraceOut_analogValues_12[0] := Binding_0_analogValues[12];
   TraceOut_analogValues_13[0] := Binding_0_analogValues[13];
   TraceOut_analogValues_14[0] := Binding_0_analogValues[14];
   TraceOut_channels_1_enable[0] := Binding_0_channels[1].enable;
   TraceOut_channels_1_hiLIM[0] := Binding_0_channels[1].hiLIM;
   TraceOut_channels_1_loLIM[0] := Binding_0_channels[1].loLIM;
   TraceOut_channels_1_bipolar[0] := Binding_0_channels[1].bipolar;
   TraceOut_channels_1_measuringMode[0] := Binding_0_channels[1].measuringMode;
   TraceOut_channels_1_retVal[0] := Binding_0_channels[1].retVal;
   TraceOut_channels_1_outputValue[0] := Binding_0_channels[1].outputValue;
   TraceOut_channels_2_enable[0] := Binding_0_channels[2].enable;
   TraceOut_channels_2_hiLIM[0] := Binding_0_channels[2].hiLIM;
   TraceOut_channels_2_loLIM[0] := Binding_0_channels[2].loLIM;
   TraceOut_channels_2_bipolar[0] := Binding_0_channels[2].bipolar;
   TraceOut_channels_2_measuringMode[0] := Binding_0_channels[2].measuringMode;
   TraceOut_channels_2_retVal[0] := Binding_0_channels[2].retVal;
   TraceOut_channels_2_outputValue[0] := Binding_0_channels[2].outputValue;
   TraceOut_channels_3_enable[0] := Binding_0_channels[3].enable;
   TraceOut_channels_3_hiLIM[0] := Binding_0_channels[3].hiLIM;
   TraceOut_channels_3_loLIM[0] := Binding_0_channels[3].loLIM;
   TraceOut_channels_3_bipolar[0] := Binding_0_channels[3].bipolar;
   TraceOut_channels_3_measuringMode[0] := Binding_0_channels[3].measuringMode;
   TraceOut_channels_3_retVal[0] := Binding_0_channels[3].retVal;
   TraceOut_channels_3_outputValue[0] := Binding_0_channels[3].outputValue;
   TraceOut_channels_4_enable[0] := Binding_0_channels[4].enable;
   TraceOut_channels_4_hiLIM[0] := Binding_0_channels[4].hiLIM;
   TraceOut_channels_4_loLIM[0] := Binding_0_channels[4].loLIM;
   TraceOut_channels_4_bipolar[0] := Binding_0_channels[4].bipolar;
   TraceOut_channels_4_measuringMode[0] := Binding_0_channels[4].measuringMode;
   TraceOut_channels_4_retVal[0] := Binding_0_channels[4].retVal;
   TraceOut_channels_4_outputValue[0] := Binding_0_channels[4].outputValue;
   TraceOut_channels_5_enable[0] := Binding_0_channels[5].enable;
   TraceOut_channels_5_hiLIM[0] := Binding_0_channels[5].hiLIM;
   TraceOut_channels_5_loLIM[0] := Binding_0_channels[5].loLIM;
   TraceOut_channels_5_bipolar[0] := Binding_0_channels[5].bipolar;
   TraceOut_channels_5_measuringMode[0] := Binding_0_channels[5].measuringMode;
   TraceOut_channels_5_retVal[0] := Binding_0_channels[5].retVal;
   TraceOut_channels_5_outputValue[0] := Binding_0_channels[5].outputValue;
   TraceOut_channels_6_enable[0] := Binding_0_channels[6].enable;
   TraceOut_channels_6_hiLIM[0] := Binding_0_channels[6].hiLIM;
   TraceOut_channels_6_loLIM[0] := Binding_0_channels[6].loLIM;
   TraceOut_channels_6_bipolar[0] := Binding_0_channels[6].bipolar;
   TraceOut_channels_6_measuringMode[0] := Binding_0_channels[6].measuringMode;
   TraceOut_channels_6_retVal[0] := Binding_0_channels[6].retVal;
   TraceOut_channels_6_outputValue[0] := Binding_0_channels[6].outputValue;
   TraceOut_channels_7_enable[0] := Binding_0_channels[7].enable;
   TraceOut_channels_7_hiLIM[0] := Binding_0_channels[7].hiLIM;
   TraceOut_channels_7_loLIM[0] := Binding_0_channels[7].loLIM;
   TraceOut_channels_7_bipolar[0] := Binding_0_channels[7].bipolar;
   TraceOut_channels_7_measuringMode[0] := Binding_0_channels[7].measuringMode;
   TraceOut_channels_7_retVal[0] := Binding_0_channels[7].retVal;
   TraceOut_channels_7_outputValue[0] := Binding_0_channels[7].outputValue;
   TraceOut_channels_8_enable[0] := Binding_0_channels[8].enable;
   TraceOut_channels_8_hiLIM[0] := Binding_0_channels[8].hiLIM;
   TraceOut_channels_8_loLIM[0] := Binding_0_channels[8].loLIM;
   TraceOut_channels_8_bipolar[0] := Binding_0_channels[8].bipolar;
   TraceOut_channels_8_measuringMode[0] := Binding_0_channels[8].measuringMode;
   TraceOut_channels_8_retVal[0] := Binding_0_channels[8].retVal;
   TraceOut_channels_8_outputValue[0] := Binding_0_channels[8].outputValue;
   TraceOut_channels_9_enable[0] := Binding_0_channels[9].enable;
   TraceOut_channels_9_hiLIM[0] := Binding_0_channels[9].hiLIM;
   TraceOut_channels_9_loLIM[0] := Binding_0_channels[9].loLIM;
   TraceOut_channels_9_bipolar[0] := Binding_0_channels[9].bipolar;
   TraceOut_channels_9_measuringMode[0] := Binding_0_channels[9].measuringMode;
   TraceOut_channels_9_retVal[0] := Binding_0_channels[9].retVal;
   TraceOut_channels_9_outputValue[0] := Binding_0_channels[9].outputValue;
   TraceOut_channels_10_enable[0] := Binding_0_channels[10].enable;
   TraceOut_channels_10_hiLIM[0] := Binding_0_channels[10].hiLIM;
   TraceOut_channels_10_loLIM[0] := Binding_0_channels[10].loLIM;
   TraceOut_channels_10_bipolar[0] := Binding_0_channels[10].bipolar;
   TraceOut_channels_10_measuringMode[0] := Binding_0_channels[10].measuringMode;
   TraceOut_channels_10_retVal[0] := Binding_0_channels[10].retVal;
   TraceOut_channels_10_outputValue[0] := Binding_0_channels[10].outputValue;
   TraceOut_channels_11_enable[0] := Binding_0_channels[11].enable;
   TraceOut_channels_11_hiLIM[0] := Binding_0_channels[11].hiLIM;
   TraceOut_channels_11_loLIM[0] := Binding_0_channels[11].loLIM;
   TraceOut_channels_11_bipolar[0] := Binding_0_channels[11].bipolar;
   TraceOut_channels_11_measuringMode[0] := Binding_0_channels[11].measuringMode;
   TraceOut_channels_11_retVal[0] := Binding_0_channels[11].retVal;
   TraceOut_channels_11_outputValue[0] := Binding_0_channels[11].outputValue;
   TraceOut_channels_12_enable[0] := Binding_0_channels[12].enable;
   TraceOut_channels_12_hiLIM[0] := Binding_0_channels[12].hiLIM;
   TraceOut_channels_12_loLIM[0] := Binding_0_channels[12].loLIM;
   TraceOut_channels_12_bipolar[0] := Binding_0_channels[12].bipolar;
   TraceOut_channels_12_measuringMode[0] := Binding_0_channels[12].measuringMode;
   TraceOut_channels_12_retVal[0] := Binding_0_channels[12].retVal;
   TraceOut_channels_12_outputValue[0] := Binding_0_channels[12].outputValue;
   TraceOut_channels_13_enable[0] := Binding_0_channels[13].enable;
   TraceOut_channels_13_hiLIM[0] := Binding_0_channels[13].hiLIM;
   TraceOut_channels_13_loLIM[0] := Binding_0_channels[13].loLIM;
   TraceOut_channels_13_bipolar[0] := Binding_0_channels[13].bipolar;
   TraceOut_channels_13_measuringMode[0] := Binding_0_channels[13].measuringMode;
   TraceOut_channels_13_retVal[0] := Binding_0_channels[13].retVal;
   TraceOut_channels_13_outputValue[0] := Binding_0_channels[13].outputValue;
   TraceOut_channels_14_enable[0] := Binding_0_channels[14].enable;
   TraceOut_channels_14_hiLIM[0] := Binding_0_channels[14].hiLIM;
   TraceOut_channels_14_loLIM[0] := Binding_0_channels[14].loLIM;
   TraceOut_channels_14_bipolar[0] := Binding_0_channels[14].bipolar;
   TraceOut_channels_14_measuringMode[0] := Binding_0_channels[14].measuringMode;
   TraceOut_channels_14_retVal[0] := Binding_0_channels[14].retVal;
   TraceOut_channels_14_outputValue[0] := Binding_0_channels[14].outputValue;
   BenchCalls := BenchCalls + 1;
 1:
   Binding_1_analogValues[1] := INT#32767;
   Binding_1_analogValues[2] := INT#-32768;
   Binding_1_analogValues[3] := INT#32767;
   Binding_1_analogValues[4] := INT#100;
   Binding_1_analogValues[5] := INT#-101;
   Binding_1_analogValues[6] := INT#500;
   Binding_1_analogValues[7] := INT#27648;
   Binding_1_analogValues[8] := INT#-27648;
   Binding_1_analogValues[9] := INT#13824;
   Binding_1_analogValues[10] := INT#777;
   Binding_1_channels[1].enable := TRUE;
   Binding_1_channels[1].hiLIM := REAL#27648.0;
   Binding_1_channels[1].loLIM := REAL#0.0;
   Binding_1_channels[1].bipolar := FALSE;
   Binding_1_channels[1].measuringMode := INT#0;
   Binding_1_channels[1].retVal := WORD#31;
   Binding_1_channels[1].outputValue := REAL#-1.0;
   Binding_1_channels[2].enable := TRUE;
   Binding_1_channels[2].hiLIM := REAL#27648.0;
   Binding_1_channels[2].loLIM := REAL#-27648.0;
   Binding_1_channels[2].bipolar := TRUE;
   Binding_1_channels[2].measuringMode := INT#0;
   Binding_1_channels[2].retVal := WORD#32;
   Binding_1_channels[2].outputValue := REAL#-2.0;
   Binding_1_channels[3].enable := TRUE;
   Binding_1_channels[3].hiLIM := REAL#27648.0;
   Binding_1_channels[3].loLIM := REAL#-27648.0;
   Binding_1_channels[3].bipolar := TRUE;
   Binding_1_channels[3].measuringMode := INT#0;
   Binding_1_channels[3].retVal := WORD#33;
   Binding_1_channels[3].outputValue := REAL#-3.0;
   Binding_1_channels[4].enable := TRUE;
   Binding_1_channels[4].hiLIM := REAL#0.0;
   Binding_1_channels[4].loLIM := REAL#0.0;
   Binding_1_channels[4].bipolar := FALSE;
   Binding_1_channels[4].measuringMode := INT#-1;
   Binding_1_channels[4].retVal := WORD#34;
   Binding_1_channels[4].outputValue := REAL#-4.0;
   Binding_1_channels[5].enable := TRUE;
   Binding_1_channels[5].hiLIM := REAL#-1.0;
   Binding_1_channels[5].loLIM := REAL#1.0;
   Binding_1_channels[5].bipolar := TRUE;
   Binding_1_channels[5].measuringMode := INT#3;
   Binding_1_channels[5].retVal := WORD#35;
   Binding_1_channels[5].outputValue := REAL#-5.0;
   Binding_1_channels[6].enable := TRUE;
   Binding_1_channels[6].hiLIM := REAL#5.0;
   Binding_1_channels[6].loLIM := REAL#5.0;
   Binding_1_channels[6].bipolar := FALSE;
   Binding_1_channels[6].measuringMode := INT#1;
   Binding_1_channels[6].retVal := WORD#36;
   Binding_1_channels[6].outputValue := REAL#-6.0;
   Binding_1_channels[7].enable := TRUE;
   Binding_1_channels[7].hiLIM := REAL#-2.0;
   Binding_1_channels[7].loLIM := REAL#2.0;
   Binding_1_channels[7].bipolar := TRUE;
   Binding_1_channels[7].measuringMode := INT#2;
   Binding_1_channels[7].retVal := WORD#37;
   Binding_1_channels[7].outputValue := REAL#-7.0;
   Binding_1_channels[8].enable := TRUE;
   Binding_1_channels[8].hiLIM := REAL#1.0;
   Binding_1_channels[8].loLIM := REAL#1.0;
   Binding_1_channels[8].bipolar := FALSE;
   Binding_1_channels[8].measuringMode := INT#0;
   Binding_1_channels[8].retVal := WORD#38;
   Binding_1_channels[8].outputValue := REAL#-8.0;
   Binding_1_channels[9].enable := FALSE;
   Binding_1_channels[9].hiLIM := REAL#-1.0;
   Binding_1_channels[9].loLIM := REAL#1.0;
   Binding_1_channels[9].bipolar := TRUE;
   Binding_1_channels[9].measuringMode := INT#99;
   Binding_1_channels[9].retVal := WORD#39;
   Binding_1_channels[9].outputValue := REAL#-9.0;
   BenchUut1.count := DINT#0;
   TraceIn_count[1] := BenchUut1.count;
   TraceInIO_analogValues_e0_INT[1] := Binding_1_analogValues[1];
   TraceInIO_analogValues_e1_INT[1] := Binding_1_analogValues[2];
   TraceInIO_analogValues_e2_INT[1] := Binding_1_analogValues[3];
   TraceInIO_analogValues_e3_INT[1] := Binding_1_analogValues[4];
   TraceInIO_analogValues_e4_INT[1] := Binding_1_analogValues[5];
   TraceInIO_analogValues_e5_INT[1] := Binding_1_analogValues[6];
   TraceInIO_analogValues_e6_INT[1] := Binding_1_analogValues[7];
   TraceInIO_analogValues_e7_INT[1] := Binding_1_analogValues[8];
   TraceInIO_analogValues_e8_INT[1] := Binding_1_analogValues[9];
   TraceInIO_analogValues_e9_INT[1] := Binding_1_analogValues[10];
   TraceInIO_channels_e0_enable_BOOL[1] := Binding_1_channels[1].enable;
   TraceInIO_channels_e0_hiLIM_REAL[1] := Binding_1_channels[1].hiLIM;
   TraceInIO_channels_e0_loLIM_REAL[1] := Binding_1_channels[1].loLIM;
   TraceInIO_channels_e0_bipolar_BOOL[1] := Binding_1_channels[1].bipolar;
   TraceInIO_channels_e0_measuringMode_INT[1] := Binding_1_channels[1].measuringMode;
   TraceInIO_channels_e0_retVal_WORD[1] := Binding_1_channels[1].retVal;
   TraceInIO_channels_e0_outputValue_REAL[1] := Binding_1_channels[1].outputValue;
   TraceInIO_channels_e1_enable_BOOL[1] := Binding_1_channels[2].enable;
   TraceInIO_channels_e1_hiLIM_REAL[1] := Binding_1_channels[2].hiLIM;
   TraceInIO_channels_e1_loLIM_REAL[1] := Binding_1_channels[2].loLIM;
   TraceInIO_channels_e1_bipolar_BOOL[1] := Binding_1_channels[2].bipolar;
   TraceInIO_channels_e1_measuringMode_INT[1] := Binding_1_channels[2].measuringMode;
   TraceInIO_channels_e1_retVal_WORD[1] := Binding_1_channels[2].retVal;
   TraceInIO_channels_e1_outputValue_REAL[1] := Binding_1_channels[2].outputValue;
   TraceInIO_channels_e2_enable_BOOL[1] := Binding_1_channels[3].enable;
   TraceInIO_channels_e2_hiLIM_REAL[1] := Binding_1_channels[3].hiLIM;
   TraceInIO_channels_e2_loLIM_REAL[1] := Binding_1_channels[3].loLIM;
   TraceInIO_channels_e2_bipolar_BOOL[1] := Binding_1_channels[3].bipolar;
   TraceInIO_channels_e2_measuringMode_INT[1] := Binding_1_channels[3].measuringMode;
   TraceInIO_channels_e2_retVal_WORD[1] := Binding_1_channels[3].retVal;
   TraceInIO_channels_e2_outputValue_REAL[1] := Binding_1_channels[3].outputValue;
   TraceInIO_channels_e3_enable_BOOL[1] := Binding_1_channels[4].enable;
   TraceInIO_channels_e3_hiLIM_REAL[1] := Binding_1_channels[4].hiLIM;
   TraceInIO_channels_e3_loLIM_REAL[1] := Binding_1_channels[4].loLIM;
   TraceInIO_channels_e3_bipolar_BOOL[1] := Binding_1_channels[4].bipolar;
   TraceInIO_channels_e3_measuringMode_INT[1] := Binding_1_channels[4].measuringMode;
   TraceInIO_channels_e3_retVal_WORD[1] := Binding_1_channels[4].retVal;
   TraceInIO_channels_e3_outputValue_REAL[1] := Binding_1_channels[4].outputValue;
   TraceInIO_channels_e4_enable_BOOL[1] := Binding_1_channels[5].enable;
   TraceInIO_channels_e4_hiLIM_REAL[1] := Binding_1_channels[5].hiLIM;
   TraceInIO_channels_e4_loLIM_REAL[1] := Binding_1_channels[5].loLIM;
   TraceInIO_channels_e4_bipolar_BOOL[1] := Binding_1_channels[5].bipolar;
   TraceInIO_channels_e4_measuringMode_INT[1] := Binding_1_channels[5].measuringMode;
   TraceInIO_channels_e4_retVal_WORD[1] := Binding_1_channels[5].retVal;
   TraceInIO_channels_e4_outputValue_REAL[1] := Binding_1_channels[5].outputValue;
   TraceInIO_channels_e5_enable_BOOL[1] := Binding_1_channels[6].enable;
   TraceInIO_channels_e5_hiLIM_REAL[1] := Binding_1_channels[6].hiLIM;
   TraceInIO_channels_e5_loLIM_REAL[1] := Binding_1_channels[6].loLIM;
   TraceInIO_channels_e5_bipolar_BOOL[1] := Binding_1_channels[6].bipolar;
   TraceInIO_channels_e5_measuringMode_INT[1] := Binding_1_channels[6].measuringMode;
   TraceInIO_channels_e5_retVal_WORD[1] := Binding_1_channels[6].retVal;
   TraceInIO_channels_e5_outputValue_REAL[1] := Binding_1_channels[6].outputValue;
   TraceInIO_channels_e6_enable_BOOL[1] := Binding_1_channels[7].enable;
   TraceInIO_channels_e6_hiLIM_REAL[1] := Binding_1_channels[7].hiLIM;
   TraceInIO_channels_e6_loLIM_REAL[1] := Binding_1_channels[7].loLIM;
   TraceInIO_channels_e6_bipolar_BOOL[1] := Binding_1_channels[7].bipolar;
   TraceInIO_channels_e6_measuringMode_INT[1] := Binding_1_channels[7].measuringMode;
   TraceInIO_channels_e6_retVal_WORD[1] := Binding_1_channels[7].retVal;
   TraceInIO_channels_e6_outputValue_REAL[1] := Binding_1_channels[7].outputValue;
   TraceInIO_channels_e7_enable_BOOL[1] := Binding_1_channels[8].enable;
   TraceInIO_channels_e7_hiLIM_REAL[1] := Binding_1_channels[8].hiLIM;
   TraceInIO_channels_e7_loLIM_REAL[1] := Binding_1_channels[8].loLIM;
   TraceInIO_channels_e7_bipolar_BOOL[1] := Binding_1_channels[8].bipolar;
   TraceInIO_channels_e7_measuringMode_INT[1] := Binding_1_channels[8].measuringMode;
   TraceInIO_channels_e7_retVal_WORD[1] := Binding_1_channels[8].retVal;
   TraceInIO_channels_e7_outputValue_REAL[1] := Binding_1_channels[8].outputValue;
   TraceInIO_channels_e8_enable_BOOL[1] := Binding_1_channels[9].enable;
   TraceInIO_channels_e8_hiLIM_REAL[1] := Binding_1_channels[9].hiLIM;
   TraceInIO_channels_e8_loLIM_REAL[1] := Binding_1_channels[9].loLIM;
   TraceInIO_channels_e8_bipolar_BOOL[1] := Binding_1_channels[9].bipolar;
   TraceInIO_channels_e8_measuringMode_INT[1] := Binding_1_channels[9].measuringMode;
   TraceInIO_channels_e8_retVal_WORD[1] := Binding_1_channels[9].retVal;
   TraceInIO_channels_e8_outputValue_REAL[1] := Binding_1_channels[9].outputValue;
   BenchUut1(analogValues := Binding_1_analogValues, channels := Binding_1_channels);
   TraceOut_analogValues_1[1] := Binding_1_analogValues[1];
   TraceOut_analogValues_2[1] := Binding_1_analogValues[2];
   TraceOut_analogValues_3[1] := Binding_1_analogValues[3];
   TraceOut_analogValues_4[1] := Binding_1_analogValues[4];
   TraceOut_analogValues_5[1] := Binding_1_analogValues[5];
   TraceOut_analogValues_6[1] := Binding_1_analogValues[6];
   TraceOut_analogValues_7[1] := Binding_1_analogValues[7];
   TraceOut_analogValues_8[1] := Binding_1_analogValues[8];
   TraceOut_analogValues_9[1] := Binding_1_analogValues[9];
   TraceOut_analogValues_10[1] := Binding_1_analogValues[10];
   TraceOut_channels_1_enable[1] := Binding_1_channels[1].enable;
   TraceOut_channels_1_hiLIM[1] := Binding_1_channels[1].hiLIM;
   TraceOut_channels_1_loLIM[1] := Binding_1_channels[1].loLIM;
   TraceOut_channels_1_bipolar[1] := Binding_1_channels[1].bipolar;
   TraceOut_channels_1_measuringMode[1] := Binding_1_channels[1].measuringMode;
   TraceOut_channels_1_retVal[1] := Binding_1_channels[1].retVal;
   TraceOut_channels_1_outputValue[1] := Binding_1_channels[1].outputValue;
   TraceOut_channels_2_enable[1] := Binding_1_channels[2].enable;
   TraceOut_channels_2_hiLIM[1] := Binding_1_channels[2].hiLIM;
   TraceOut_channels_2_loLIM[1] := Binding_1_channels[2].loLIM;
   TraceOut_channels_2_bipolar[1] := Binding_1_channels[2].bipolar;
   TraceOut_channels_2_measuringMode[1] := Binding_1_channels[2].measuringMode;
   TraceOut_channels_2_retVal[1] := Binding_1_channels[2].retVal;
   TraceOut_channels_2_outputValue[1] := Binding_1_channels[2].outputValue;
   TraceOut_channels_3_enable[1] := Binding_1_channels[3].enable;
   TraceOut_channels_3_hiLIM[1] := Binding_1_channels[3].hiLIM;
   TraceOut_channels_3_loLIM[1] := Binding_1_channels[3].loLIM;
   TraceOut_channels_3_bipolar[1] := Binding_1_channels[3].bipolar;
   TraceOut_channels_3_measuringMode[1] := Binding_1_channels[3].measuringMode;
   TraceOut_channels_3_retVal[1] := Binding_1_channels[3].retVal;
   TraceOut_channels_3_outputValue[1] := Binding_1_channels[3].outputValue;
   TraceOut_channels_4_enable[1] := Binding_1_channels[4].enable;
   TraceOut_channels_4_hiLIM[1] := Binding_1_channels[4].hiLIM;
   TraceOut_channels_4_loLIM[1] := Binding_1_channels[4].loLIM;
   TraceOut_channels_4_bipolar[1] := Binding_1_channels[4].bipolar;
   TraceOut_channels_4_measuringMode[1] := Binding_1_channels[4].measuringMode;
   TraceOut_channels_4_retVal[1] := Binding_1_channels[4].retVal;
   TraceOut_channels_4_outputValue[1] := Binding_1_channels[4].outputValue;
   TraceOut_channels_5_enable[1] := Binding_1_channels[5].enable;
   TraceOut_channels_5_hiLIM[1] := Binding_1_channels[5].hiLIM;
   TraceOut_channels_5_loLIM[1] := Binding_1_channels[5].loLIM;
   TraceOut_channels_5_bipolar[1] := Binding_1_channels[5].bipolar;
   TraceOut_channels_5_measuringMode[1] := Binding_1_channels[5].measuringMode;
   TraceOut_channels_5_retVal[1] := Binding_1_channels[5].retVal;
   TraceOut_channels_5_outputValue[1] := Binding_1_channels[5].outputValue;
   TraceOut_channels_6_enable[1] := Binding_1_channels[6].enable;
   TraceOut_channels_6_hiLIM[1] := Binding_1_channels[6].hiLIM;
   TraceOut_channels_6_loLIM[1] := Binding_1_channels[6].loLIM;
   TraceOut_channels_6_bipolar[1] := Binding_1_channels[6].bipolar;
   TraceOut_channels_6_measuringMode[1] := Binding_1_channels[6].measuringMode;
   TraceOut_channels_6_retVal[1] := Binding_1_channels[6].retVal;
   TraceOut_channels_6_outputValue[1] := Binding_1_channels[6].outputValue;
   TraceOut_channels_7_enable[1] := Binding_1_channels[7].enable;
   TraceOut_channels_7_hiLIM[1] := Binding_1_channels[7].hiLIM;
   TraceOut_channels_7_loLIM[1] := Binding_1_channels[7].loLIM;
   TraceOut_channels_7_bipolar[1] := Binding_1_channels[7].bipolar;
   TraceOut_channels_7_measuringMode[1] := Binding_1_channels[7].measuringMode;
   TraceOut_channels_7_retVal[1] := Binding_1_channels[7].retVal;
   TraceOut_channels_7_outputValue[1] := Binding_1_channels[7].outputValue;
   TraceOut_channels_8_enable[1] := Binding_1_channels[8].enable;
   TraceOut_channels_8_hiLIM[1] := Binding_1_channels[8].hiLIM;
   TraceOut_channels_8_loLIM[1] := Binding_1_channels[8].loLIM;
   TraceOut_channels_8_bipolar[1] := Binding_1_channels[8].bipolar;
   TraceOut_channels_8_measuringMode[1] := Binding_1_channels[8].measuringMode;
   TraceOut_channels_8_retVal[1] := Binding_1_channels[8].retVal;
   TraceOut_channels_8_outputValue[1] := Binding_1_channels[8].outputValue;
   TraceOut_channels_9_enable[1] := Binding_1_channels[9].enable;
   TraceOut_channels_9_hiLIM[1] := Binding_1_channels[9].hiLIM;
   TraceOut_channels_9_loLIM[1] := Binding_1_channels[9].loLIM;
   TraceOut_channels_9_bipolar[1] := Binding_1_channels[9].bipolar;
   TraceOut_channels_9_measuringMode[1] := Binding_1_channels[9].measuringMode;
   TraceOut_channels_9_retVal[1] := Binding_1_channels[9].retVal;
   TraceOut_channels_9_outputValue[1] := Binding_1_channels[9].outputValue;
   BenchCalls := BenchCalls + 1;
 2:
   Binding_1_analogValues[1] := INT#32767;
   Binding_1_analogValues[2] := INT#-32768;
   Binding_1_analogValues[3] := INT#32767;
   Binding_1_analogValues[4] := INT#100;
   Binding_1_analogValues[5] := INT#-101;
   Binding_1_analogValues[6] := INT#500;
   Binding_1_analogValues[7] := INT#27648;
   Binding_1_analogValues[8] := INT#-27648;
   Binding_1_analogValues[9] := INT#13824;
   Binding_1_analogValues[10] := INT#777;
   Binding_1_channels[1].enable := TRUE;
   Binding_1_channels[1].hiLIM := REAL#27648.0;
   Binding_1_channels[1].loLIM := REAL#0.0;
   Binding_1_channels[1].bipolar := FALSE;
   Binding_1_channels[1].measuringMode := INT#0;
   Binding_1_channels[1].retVal := WORD#31;
   Binding_1_channels[1].outputValue := REAL#-1.0;
   Binding_1_channels[2].enable := TRUE;
   Binding_1_channels[2].hiLIM := REAL#27648.0;
   Binding_1_channels[2].loLIM := REAL#-27648.0;
   Binding_1_channels[2].bipolar := TRUE;
   Binding_1_channels[2].measuringMode := INT#0;
   Binding_1_channels[2].retVal := WORD#32;
   Binding_1_channels[2].outputValue := REAL#-2.0;
   Binding_1_channels[3].enable := TRUE;
   Binding_1_channels[3].hiLIM := REAL#27648.0;
   Binding_1_channels[3].loLIM := REAL#-27648.0;
   Binding_1_channels[3].bipolar := TRUE;
   Binding_1_channels[3].measuringMode := INT#0;
   Binding_1_channels[3].retVal := WORD#33;
   Binding_1_channels[3].outputValue := REAL#-3.0;
   Binding_1_channels[4].enable := TRUE;
   Binding_1_channels[4].hiLIM := REAL#0.0;
   Binding_1_channels[4].loLIM := REAL#0.0;
   Binding_1_channels[4].bipolar := FALSE;
   Binding_1_channels[4].measuringMode := INT#-1;
   Binding_1_channels[4].retVal := WORD#34;
   Binding_1_channels[4].outputValue := REAL#-4.0;
   Binding_1_channels[5].enable := TRUE;
   Binding_1_channels[5].hiLIM := REAL#-1.0;
   Binding_1_channels[5].loLIM := REAL#1.0;
   Binding_1_channels[5].bipolar := TRUE;
   Binding_1_channels[5].measuringMode := INT#3;
   Binding_1_channels[5].retVal := WORD#35;
   Binding_1_channels[5].outputValue := REAL#-5.0;
   Binding_1_channels[6].enable := TRUE;
   Binding_1_channels[6].hiLIM := REAL#5.0;
   Binding_1_channels[6].loLIM := REAL#5.0;
   Binding_1_channels[6].bipolar := FALSE;
   Binding_1_channels[6].measuringMode := INT#1;
   Binding_1_channels[6].retVal := WORD#36;
   Binding_1_channels[6].outputValue := REAL#-6.0;
   Binding_1_channels[7].enable := TRUE;
   Binding_1_channels[7].hiLIM := REAL#-2.0;
   Binding_1_channels[7].loLIM := REAL#2.0;
   Binding_1_channels[7].bipolar := TRUE;
   Binding_1_channels[7].measuringMode := INT#2;
   Binding_1_channels[7].retVal := WORD#37;
   Binding_1_channels[7].outputValue := REAL#-7.0;
   Binding_1_channels[8].enable := TRUE;
   Binding_1_channels[8].hiLIM := REAL#1.0;
   Binding_1_channels[8].loLIM := REAL#1.0;
   Binding_1_channels[8].bipolar := FALSE;
   Binding_1_channels[8].measuringMode := INT#0;
   Binding_1_channels[8].retVal := WORD#38;
   Binding_1_channels[8].outputValue := REAL#-8.0;
   Binding_1_channels[9].enable := FALSE;
   Binding_1_channels[9].hiLIM := REAL#-1.0;
   Binding_1_channels[9].loLIM := REAL#1.0;
   Binding_1_channels[9].bipolar := TRUE;
   Binding_1_channels[9].measuringMode := INT#99;
   Binding_1_channels[9].retVal := WORD#39;
   Binding_1_channels[9].outputValue := REAL#-9.0;
   BenchUut1.count := DINT#9;
   TraceIn_count[2] := BenchUut1.count;
   TraceInIO_analogValues_e0_INT[2] := Binding_1_analogValues[1];
   TraceInIO_analogValues_e1_INT[2] := Binding_1_analogValues[2];
   TraceInIO_analogValues_e2_INT[2] := Binding_1_analogValues[3];
   TraceInIO_analogValues_e3_INT[2] := Binding_1_analogValues[4];
   TraceInIO_analogValues_e4_INT[2] := Binding_1_analogValues[5];
   TraceInIO_analogValues_e5_INT[2] := Binding_1_analogValues[6];
   TraceInIO_analogValues_e6_INT[2] := Binding_1_analogValues[7];
   TraceInIO_analogValues_e7_INT[2] := Binding_1_analogValues[8];
   TraceInIO_analogValues_e8_INT[2] := Binding_1_analogValues[9];
   TraceInIO_analogValues_e9_INT[2] := Binding_1_analogValues[10];
   TraceInIO_channels_e0_enable_BOOL[2] := Binding_1_channels[1].enable;
   TraceInIO_channels_e0_hiLIM_REAL[2] := Binding_1_channels[1].hiLIM;
   TraceInIO_channels_e0_loLIM_REAL[2] := Binding_1_channels[1].loLIM;
   TraceInIO_channels_e0_bipolar_BOOL[2] := Binding_1_channels[1].bipolar;
   TraceInIO_channels_e0_measuringMode_INT[2] := Binding_1_channels[1].measuringMode;
   TraceInIO_channels_e0_retVal_WORD[2] := Binding_1_channels[1].retVal;
   TraceInIO_channels_e0_outputValue_REAL[2] := Binding_1_channels[1].outputValue;
   TraceInIO_channels_e1_enable_BOOL[2] := Binding_1_channels[2].enable;
   TraceInIO_channels_e1_hiLIM_REAL[2] := Binding_1_channels[2].hiLIM;
   TraceInIO_channels_e1_loLIM_REAL[2] := Binding_1_channels[2].loLIM;
   TraceInIO_channels_e1_bipolar_BOOL[2] := Binding_1_channels[2].bipolar;
   TraceInIO_channels_e1_measuringMode_INT[2] := Binding_1_channels[2].measuringMode;
   TraceInIO_channels_e1_retVal_WORD[2] := Binding_1_channels[2].retVal;
   TraceInIO_channels_e1_outputValue_REAL[2] := Binding_1_channels[2].outputValue;
   TraceInIO_channels_e2_enable_BOOL[2] := Binding_1_channels[3].enable;
   TraceInIO_channels_e2_hiLIM_REAL[2] := Binding_1_channels[3].hiLIM;
   TraceInIO_channels_e2_loLIM_REAL[2] := Binding_1_channels[3].loLIM;
   TraceInIO_channels_e2_bipolar_BOOL[2] := Binding_1_channels[3].bipolar;
   TraceInIO_channels_e2_measuringMode_INT[2] := Binding_1_channels[3].measuringMode;
   TraceInIO_channels_e2_retVal_WORD[2] := Binding_1_channels[3].retVal;
   TraceInIO_channels_e2_outputValue_REAL[2] := Binding_1_channels[3].outputValue;
   TraceInIO_channels_e3_enable_BOOL[2] := Binding_1_channels[4].enable;
   TraceInIO_channels_e3_hiLIM_REAL[2] := Binding_1_channels[4].hiLIM;
   TraceInIO_channels_e3_loLIM_REAL[2] := Binding_1_channels[4].loLIM;
   TraceInIO_channels_e3_bipolar_BOOL[2] := Binding_1_channels[4].bipolar;
   TraceInIO_channels_e3_measuringMode_INT[2] := Binding_1_channels[4].measuringMode;
   TraceInIO_channels_e3_retVal_WORD[2] := Binding_1_channels[4].retVal;
   TraceInIO_channels_e3_outputValue_REAL[2] := Binding_1_channels[4].outputValue;
   TraceInIO_channels_e4_enable_BOOL[2] := Binding_1_channels[5].enable;
   TraceInIO_channels_e4_hiLIM_REAL[2] := Binding_1_channels[5].hiLIM;
   TraceInIO_channels_e4_loLIM_REAL[2] := Binding_1_channels[5].loLIM;
   TraceInIO_channels_e4_bipolar_BOOL[2] := Binding_1_channels[5].bipolar;
   TraceInIO_channels_e4_measuringMode_INT[2] := Binding_1_channels[5].measuringMode;
   TraceInIO_channels_e4_retVal_WORD[2] := Binding_1_channels[5].retVal;
   TraceInIO_channels_e4_outputValue_REAL[2] := Binding_1_channels[5].outputValue;
   TraceInIO_channels_e5_enable_BOOL[2] := Binding_1_channels[6].enable;
   TraceInIO_channels_e5_hiLIM_REAL[2] := Binding_1_channels[6].hiLIM;
   TraceInIO_channels_e5_loLIM_REAL[2] := Binding_1_channels[6].loLIM;
   TraceInIO_channels_e5_bipolar_BOOL[2] := Binding_1_channels[6].bipolar;
   TraceInIO_channels_e5_measuringMode_INT[2] := Binding_1_channels[6].measuringMode;
   TraceInIO_channels_e5_retVal_WORD[2] := Binding_1_channels[6].retVal;
   TraceInIO_channels_e5_outputValue_REAL[2] := Binding_1_channels[6].outputValue;
   TraceInIO_channels_e6_enable_BOOL[2] := Binding_1_channels[7].enable;
   TraceInIO_channels_e6_hiLIM_REAL[2] := Binding_1_channels[7].hiLIM;
   TraceInIO_channels_e6_loLIM_REAL[2] := Binding_1_channels[7].loLIM;
   TraceInIO_channels_e6_bipolar_BOOL[2] := Binding_1_channels[7].bipolar;
   TraceInIO_channels_e6_measuringMode_INT[2] := Binding_1_channels[7].measuringMode;
   TraceInIO_channels_e6_retVal_WORD[2] := Binding_1_channels[7].retVal;
   TraceInIO_channels_e6_outputValue_REAL[2] := Binding_1_channels[7].outputValue;
   TraceInIO_channels_e7_enable_BOOL[2] := Binding_1_channels[8].enable;
   TraceInIO_channels_e7_hiLIM_REAL[2] := Binding_1_channels[8].hiLIM;
   TraceInIO_channels_e7_loLIM_REAL[2] := Binding_1_channels[8].loLIM;
   TraceInIO_channels_e7_bipolar_BOOL[2] := Binding_1_channels[8].bipolar;
   TraceInIO_channels_e7_measuringMode_INT[2] := Binding_1_channels[8].measuringMode;
   TraceInIO_channels_e7_retVal_WORD[2] := Binding_1_channels[8].retVal;
   TraceInIO_channels_e7_outputValue_REAL[2] := Binding_1_channels[8].outputValue;
   TraceInIO_channels_e8_enable_BOOL[2] := Binding_1_channels[9].enable;
   TraceInIO_channels_e8_hiLIM_REAL[2] := Binding_1_channels[9].hiLIM;
   TraceInIO_channels_e8_loLIM_REAL[2] := Binding_1_channels[9].loLIM;
   TraceInIO_channels_e8_bipolar_BOOL[2] := Binding_1_channels[9].bipolar;
   TraceInIO_channels_e8_measuringMode_INT[2] := Binding_1_channels[9].measuringMode;
   TraceInIO_channels_e8_retVal_WORD[2] := Binding_1_channels[9].retVal;
   TraceInIO_channels_e8_outputValue_REAL[2] := Binding_1_channels[9].outputValue;
   BenchUut1(analogValues := Binding_1_analogValues, channels := Binding_1_channels);
   TraceOut_analogValues_1[2] := Binding_1_analogValues[1];
   TraceOut_analogValues_2[2] := Binding_1_analogValues[2];
   TraceOut_analogValues_3[2] := Binding_1_analogValues[3];
   TraceOut_analogValues_4[2] := Binding_1_analogValues[4];
   TraceOut_analogValues_5[2] := Binding_1_analogValues[5];
   TraceOut_analogValues_6[2] := Binding_1_analogValues[6];
   TraceOut_analogValues_7[2] := Binding_1_analogValues[7];
   TraceOut_analogValues_8[2] := Binding_1_analogValues[8];
   TraceOut_analogValues_9[2] := Binding_1_analogValues[9];
   TraceOut_analogValues_10[2] := Binding_1_analogValues[10];
   TraceOut_channels_1_enable[2] := Binding_1_channels[1].enable;
   TraceOut_channels_1_hiLIM[2] := Binding_1_channels[1].hiLIM;
   TraceOut_channels_1_loLIM[2] := Binding_1_channels[1].loLIM;
   TraceOut_channels_1_bipolar[2] := Binding_1_channels[1].bipolar;
   TraceOut_channels_1_measuringMode[2] := Binding_1_channels[1].measuringMode;
   TraceOut_channels_1_retVal[2] := Binding_1_channels[1].retVal;
   TraceOut_channels_1_outputValue[2] := Binding_1_channels[1].outputValue;
   TraceOut_channels_2_enable[2] := Binding_1_channels[2].enable;
   TraceOut_channels_2_hiLIM[2] := Binding_1_channels[2].hiLIM;
   TraceOut_channels_2_loLIM[2] := Binding_1_channels[2].loLIM;
   TraceOut_channels_2_bipolar[2] := Binding_1_channels[2].bipolar;
   TraceOut_channels_2_measuringMode[2] := Binding_1_channels[2].measuringMode;
   TraceOut_channels_2_retVal[2] := Binding_1_channels[2].retVal;
   TraceOut_channels_2_outputValue[2] := Binding_1_channels[2].outputValue;
   TraceOut_channels_3_enable[2] := Binding_1_channels[3].enable;
   TraceOut_channels_3_hiLIM[2] := Binding_1_channels[3].hiLIM;
   TraceOut_channels_3_loLIM[2] := Binding_1_channels[3].loLIM;
   TraceOut_channels_3_bipolar[2] := Binding_1_channels[3].bipolar;
   TraceOut_channels_3_measuringMode[2] := Binding_1_channels[3].measuringMode;
   TraceOut_channels_3_retVal[2] := Binding_1_channels[3].retVal;
   TraceOut_channels_3_outputValue[2] := Binding_1_channels[3].outputValue;
   TraceOut_channels_4_enable[2] := Binding_1_channels[4].enable;
   TraceOut_channels_4_hiLIM[2] := Binding_1_channels[4].hiLIM;
   TraceOut_channels_4_loLIM[2] := Binding_1_channels[4].loLIM;
   TraceOut_channels_4_bipolar[2] := Binding_1_channels[4].bipolar;
   TraceOut_channels_4_measuringMode[2] := Binding_1_channels[4].measuringMode;
   TraceOut_channels_4_retVal[2] := Binding_1_channels[4].retVal;
   TraceOut_channels_4_outputValue[2] := Binding_1_channels[4].outputValue;
   TraceOut_channels_5_enable[2] := Binding_1_channels[5].enable;
   TraceOut_channels_5_hiLIM[2] := Binding_1_channels[5].hiLIM;
   TraceOut_channels_5_loLIM[2] := Binding_1_channels[5].loLIM;
   TraceOut_channels_5_bipolar[2] := Binding_1_channels[5].bipolar;
   TraceOut_channels_5_measuringMode[2] := Binding_1_channels[5].measuringMode;
   TraceOut_channels_5_retVal[2] := Binding_1_channels[5].retVal;
   TraceOut_channels_5_outputValue[2] := Binding_1_channels[5].outputValue;
   TraceOut_channels_6_enable[2] := Binding_1_channels[6].enable;
   TraceOut_channels_6_hiLIM[2] := Binding_1_channels[6].hiLIM;
   TraceOut_channels_6_loLIM[2] := Binding_1_channels[6].loLIM;
   TraceOut_channels_6_bipolar[2] := Binding_1_channels[6].bipolar;
   TraceOut_channels_6_measuringMode[2] := Binding_1_channels[6].measuringMode;
   TraceOut_channels_6_retVal[2] := Binding_1_channels[6].retVal;
   TraceOut_channels_6_outputValue[2] := Binding_1_channels[6].outputValue;
   TraceOut_channels_7_enable[2] := Binding_1_channels[7].enable;
   TraceOut_channels_7_hiLIM[2] := Binding_1_channels[7].hiLIM;
   TraceOut_channels_7_loLIM[2] := Binding_1_channels[7].loLIM;
   TraceOut_channels_7_bipolar[2] := Binding_1_channels[7].bipolar;
   TraceOut_channels_7_measuringMode[2] := Binding_1_channels[7].measuringMode;
   TraceOut_channels_7_retVal[2] := Binding_1_channels[7].retVal;
   TraceOut_channels_7_outputValue[2] := Binding_1_channels[7].outputValue;
   TraceOut_channels_8_enable[2] := Binding_1_channels[8].enable;
   TraceOut_channels_8_hiLIM[2] := Binding_1_channels[8].hiLIM;
   TraceOut_channels_8_loLIM[2] := Binding_1_channels[8].loLIM;
   TraceOut_channels_8_bipolar[2] := Binding_1_channels[8].bipolar;
   TraceOut_channels_8_measuringMode[2] := Binding_1_channels[8].measuringMode;
   TraceOut_channels_8_retVal[2] := Binding_1_channels[8].retVal;
   TraceOut_channels_8_outputValue[2] := Binding_1_channels[8].outputValue;
   TraceOut_channels_9_enable[2] := Binding_1_channels[9].enable;
   TraceOut_channels_9_hiLIM[2] := Binding_1_channels[9].hiLIM;
   TraceOut_channels_9_loLIM[2] := Binding_1_channels[9].loLIM;
   TraceOut_channels_9_bipolar[2] := Binding_1_channels[9].bipolar;
   TraceOut_channels_9_measuringMode[2] := Binding_1_channels[9].measuringMode;
   TraceOut_channels_9_retVal[2] := Binding_1_channels[9].retVal;
   TraceOut_channels_9_outputValue[2] := Binding_1_channels[9].outputValue;
   BenchCalls := BenchCalls + 1;
 3:
   Binding_1_analogValues[1] := INT#0;
   Binding_1_analogValues[2] := INT#0;
   Binding_1_analogValues[3] := INT#0;
   Binding_1_analogValues[4] := INT#-101;
   Binding_1_analogValues[5] := INT#105;
   Binding_1_analogValues[6] := INT#1;
   Binding_1_analogValues[7] := INT#-1;
   Binding_1_analogValues[8] := INT#13824;
   Binding_1_analogValues[9] := INT#0;
   Binding_1_analogValues[10] := INT#777;
   Binding_1_channels[1].enable := FALSE;
   Binding_1_channels[1].hiLIM := REAL#27648.0;
   Binding_1_channels[1].loLIM := REAL#0.0;
   Binding_1_channels[1].bipolar := FALSE;
   Binding_1_channels[1].measuringMode := INT#0;
   Binding_1_channels[1].retVal := WORD#0;
   Binding_1_channels[1].outputValue := REAL#32767.0;
   Binding_1_channels[2].enable := TRUE;
   Binding_1_channels[2].hiLIM := REAL#27648.0;
   Binding_1_channels[2].loLIM := REAL#-27648.0;
   Binding_1_channels[2].bipolar := TRUE;
   Binding_1_channels[2].measuringMode := INT#-32768;
   Binding_1_channels[2].retVal := WORD#0;
   Binding_1_channels[2].outputValue := REAL#-32768.0;
   Binding_1_channels[3].enable := TRUE;
   Binding_1_channels[3].hiLIM := REAL#5.0;
   Binding_1_channels[3].loLIM := REAL#5.0;
   Binding_1_channels[3].bipolar := TRUE;
   Binding_1_channels[3].measuringMode := INT#0;
   Binding_1_channels[3].retVal := WORD#0;
   Binding_1_channels[3].outputValue := REAL#32767.0;
   Binding_1_channels[4].enable := TRUE;
   Binding_1_channels[4].hiLIM := REAL#10.0;
   Binding_1_channels[4].loLIM := REAL#-10.0;
   Binding_1_channels[4].bipolar := FALSE;
   Binding_1_channels[4].measuringMode := INT#1;
   Binding_1_channels[4].retVal := WORD#32769;
   Binding_1_channels[4].outputValue := REAL#-4.0;
   Binding_1_channels[5].enable := TRUE;
   Binding_1_channels[5].hiLIM := REAL#10.0;
   Binding_1_channels[5].loLIM := REAL#-10.0;
   Binding_1_channels[5].bipolar := TRUE;
   Binding_1_channels[5].measuringMode := INT#2;
   Binding_1_channels[5].retVal := WORD#32769;
   Binding_1_channels[5].outputValue := REAL#-5.0;
   Binding_1_channels[6].enable := TRUE;
   Binding_1_channels[6].hiLIM := REAL#10.0;
   Binding_1_channels[6].loLIM := REAL#-10.0;
   Binding_1_channels[6].bipolar := FALSE;
   Binding_1_channels[6].measuringMode := INT#1;
   Binding_1_channels[6].retVal := WORD#32770;
   Binding_1_channels[6].outputValue := REAL#-6.0;
   Binding_1_channels[7].enable := TRUE;
   Binding_1_channels[7].hiLIM := REAL#10.0;
   Binding_1_channels[7].loLIM := REAL#-10.0;
   Binding_1_channels[7].bipolar := TRUE;
   Binding_1_channels[7].measuringMode := INT#2;
   Binding_1_channels[7].retVal := WORD#32770;
   Binding_1_channels[7].outputValue := REAL#-7.0;
   Binding_1_channels[8].enable := TRUE;
   Binding_1_channels[8].hiLIM := REAL#1.0;
   Binding_1_channels[8].loLIM := REAL#-1.0;
   Binding_1_channels[8].bipolar := FALSE;
   Binding_1_channels[8].measuringMode := INT#0;
   Binding_1_channels[8].retVal := WORD#32770;
   Binding_1_channels[8].outputValue := REAL#-8.0;
   Binding_1_channels[9].enable := TRUE;
   Binding_1_channels[9].hiLIM := REAL#-1.0;
   Binding_1_channels[9].loLIM := REAL#1.0;
   Binding_1_channels[9].bipolar := TRUE;
   Binding_1_channels[9].measuringMode := INT#99;
   Binding_1_channels[9].retVal := WORD#39;
   Binding_1_channels[9].outputValue := REAL#-9.0;
   BenchUut1.count := DINT#9;
   TraceIn_count[3] := BenchUut1.count;
   TraceInIO_analogValues_e0_INT[3] := Binding_1_analogValues[1];
   TraceInIO_analogValues_e1_INT[3] := Binding_1_analogValues[2];
   TraceInIO_analogValues_e2_INT[3] := Binding_1_analogValues[3];
   TraceInIO_analogValues_e3_INT[3] := Binding_1_analogValues[4];
   TraceInIO_analogValues_e4_INT[3] := Binding_1_analogValues[5];
   TraceInIO_analogValues_e5_INT[3] := Binding_1_analogValues[6];
   TraceInIO_analogValues_e6_INT[3] := Binding_1_analogValues[7];
   TraceInIO_analogValues_e7_INT[3] := Binding_1_analogValues[8];
   TraceInIO_analogValues_e8_INT[3] := Binding_1_analogValues[9];
   TraceInIO_analogValues_e9_INT[3] := Binding_1_analogValues[10];
   TraceInIO_channels_e0_enable_BOOL[3] := Binding_1_channels[1].enable;
   TraceInIO_channels_e0_hiLIM_REAL[3] := Binding_1_channels[1].hiLIM;
   TraceInIO_channels_e0_loLIM_REAL[3] := Binding_1_channels[1].loLIM;
   TraceInIO_channels_e0_bipolar_BOOL[3] := Binding_1_channels[1].bipolar;
   TraceInIO_channels_e0_measuringMode_INT[3] := Binding_1_channels[1].measuringMode;
   TraceInIO_channels_e0_retVal_WORD[3] := Binding_1_channels[1].retVal;
   TraceInIO_channels_e0_outputValue_REAL[3] := Binding_1_channels[1].outputValue;
   TraceInIO_channels_e1_enable_BOOL[3] := Binding_1_channels[2].enable;
   TraceInIO_channels_e1_hiLIM_REAL[3] := Binding_1_channels[2].hiLIM;
   TraceInIO_channels_e1_loLIM_REAL[3] := Binding_1_channels[2].loLIM;
   TraceInIO_channels_e1_bipolar_BOOL[3] := Binding_1_channels[2].bipolar;
   TraceInIO_channels_e1_measuringMode_INT[3] := Binding_1_channels[2].measuringMode;
   TraceInIO_channels_e1_retVal_WORD[3] := Binding_1_channels[2].retVal;
   TraceInIO_channels_e1_outputValue_REAL[3] := Binding_1_channels[2].outputValue;
   TraceInIO_channels_e2_enable_BOOL[3] := Binding_1_channels[3].enable;
   TraceInIO_channels_e2_hiLIM_REAL[3] := Binding_1_channels[3].hiLIM;
   TraceInIO_channels_e2_loLIM_REAL[3] := Binding_1_channels[3].loLIM;
   TraceInIO_channels_e2_bipolar_BOOL[3] := Binding_1_channels[3].bipolar;
   TraceInIO_channels_e2_measuringMode_INT[3] := Binding_1_channels[3].measuringMode;
   TraceInIO_channels_e2_retVal_WORD[3] := Binding_1_channels[3].retVal;
   TraceInIO_channels_e2_outputValue_REAL[3] := Binding_1_channels[3].outputValue;
   TraceInIO_channels_e3_enable_BOOL[3] := Binding_1_channels[4].enable;
   TraceInIO_channels_e3_hiLIM_REAL[3] := Binding_1_channels[4].hiLIM;
   TraceInIO_channels_e3_loLIM_REAL[3] := Binding_1_channels[4].loLIM;
   TraceInIO_channels_e3_bipolar_BOOL[3] := Binding_1_channels[4].bipolar;
   TraceInIO_channels_e3_measuringMode_INT[3] := Binding_1_channels[4].measuringMode;
   TraceInIO_channels_e3_retVal_WORD[3] := Binding_1_channels[4].retVal;
   TraceInIO_channels_e3_outputValue_REAL[3] := Binding_1_channels[4].outputValue;
   TraceInIO_channels_e4_enable_BOOL[3] := Binding_1_channels[5].enable;
   TraceInIO_channels_e4_hiLIM_REAL[3] := Binding_1_channels[5].hiLIM;
   TraceInIO_channels_e4_loLIM_REAL[3] := Binding_1_channels[5].loLIM;
   TraceInIO_channels_e4_bipolar_BOOL[3] := Binding_1_channels[5].bipolar;
   TraceInIO_channels_e4_measuringMode_INT[3] := Binding_1_channels[5].measuringMode;
   TraceInIO_channels_e4_retVal_WORD[3] := Binding_1_channels[5].retVal;
   TraceInIO_channels_e4_outputValue_REAL[3] := Binding_1_channels[5].outputValue;
   TraceInIO_channels_e5_enable_BOOL[3] := Binding_1_channels[6].enable;
   TraceInIO_channels_e5_hiLIM_REAL[3] := Binding_1_channels[6].hiLIM;
   TraceInIO_channels_e5_loLIM_REAL[3] := Binding_1_channels[6].loLIM;
   TraceInIO_channels_e5_bipolar_BOOL[3] := Binding_1_channels[6].bipolar;
   TraceInIO_channels_e5_measuringMode_INT[3] := Binding_1_channels[6].measuringMode;
   TraceInIO_channels_e5_retVal_WORD[3] := Binding_1_channels[6].retVal;
   TraceInIO_channels_e5_outputValue_REAL[3] := Binding_1_channels[6].outputValue;
   TraceInIO_channels_e6_enable_BOOL[3] := Binding_1_channels[7].enable;
   TraceInIO_channels_e6_hiLIM_REAL[3] := Binding_1_channels[7].hiLIM;
   TraceInIO_channels_e6_loLIM_REAL[3] := Binding_1_channels[7].loLIM;
   TraceInIO_channels_e6_bipolar_BOOL[3] := Binding_1_channels[7].bipolar;
   TraceInIO_channels_e6_measuringMode_INT[3] := Binding_1_channels[7].measuringMode;
   TraceInIO_channels_e6_retVal_WORD[3] := Binding_1_channels[7].retVal;
   TraceInIO_channels_e6_outputValue_REAL[3] := Binding_1_channels[7].outputValue;
   TraceInIO_channels_e7_enable_BOOL[3] := Binding_1_channels[8].enable;
   TraceInIO_channels_e7_hiLIM_REAL[3] := Binding_1_channels[8].hiLIM;
   TraceInIO_channels_e7_loLIM_REAL[3] := Binding_1_channels[8].loLIM;
   TraceInIO_channels_e7_bipolar_BOOL[3] := Binding_1_channels[8].bipolar;
   TraceInIO_channels_e7_measuringMode_INT[3] := Binding_1_channels[8].measuringMode;
   TraceInIO_channels_e7_retVal_WORD[3] := Binding_1_channels[8].retVal;
   TraceInIO_channels_e7_outputValue_REAL[3] := Binding_1_channels[8].outputValue;
   TraceInIO_channels_e8_enable_BOOL[3] := Binding_1_channels[9].enable;
   TraceInIO_channels_e8_hiLIM_REAL[3] := Binding_1_channels[9].hiLIM;
   TraceInIO_channels_e8_loLIM_REAL[3] := Binding_1_channels[9].loLIM;
   TraceInIO_channels_e8_bipolar_BOOL[3] := Binding_1_channels[9].bipolar;
   TraceInIO_channels_e8_measuringMode_INT[3] := Binding_1_channels[9].measuringMode;
   TraceInIO_channels_e8_retVal_WORD[3] := Binding_1_channels[9].retVal;
   TraceInIO_channels_e8_outputValue_REAL[3] := Binding_1_channels[9].outputValue;
   BenchUut1(analogValues := Binding_1_analogValues, channels := Binding_1_channels);
   TraceOut_analogValues_1[3] := Binding_1_analogValues[1];
   TraceOut_analogValues_2[3] := Binding_1_analogValues[2];
   TraceOut_analogValues_3[3] := Binding_1_analogValues[3];
   TraceOut_analogValues_4[3] := Binding_1_analogValues[4];
   TraceOut_analogValues_5[3] := Binding_1_analogValues[5];
   TraceOut_analogValues_6[3] := Binding_1_analogValues[6];
   TraceOut_analogValues_7[3] := Binding_1_analogValues[7];
   TraceOut_analogValues_8[3] := Binding_1_analogValues[8];
   TraceOut_analogValues_9[3] := Binding_1_analogValues[9];
   TraceOut_analogValues_10[3] := Binding_1_analogValues[10];
   TraceOut_channels_1_enable[3] := Binding_1_channels[1].enable;
   TraceOut_channels_1_hiLIM[3] := Binding_1_channels[1].hiLIM;
   TraceOut_channels_1_loLIM[3] := Binding_1_channels[1].loLIM;
   TraceOut_channels_1_bipolar[3] := Binding_1_channels[1].bipolar;
   TraceOut_channels_1_measuringMode[3] := Binding_1_channels[1].measuringMode;
   TraceOut_channels_1_retVal[3] := Binding_1_channels[1].retVal;
   TraceOut_channels_1_outputValue[3] := Binding_1_channels[1].outputValue;
   TraceOut_channels_2_enable[3] := Binding_1_channels[2].enable;
   TraceOut_channels_2_hiLIM[3] := Binding_1_channels[2].hiLIM;
   TraceOut_channels_2_loLIM[3] := Binding_1_channels[2].loLIM;
   TraceOut_channels_2_bipolar[3] := Binding_1_channels[2].bipolar;
   TraceOut_channels_2_measuringMode[3] := Binding_1_channels[2].measuringMode;
   TraceOut_channels_2_retVal[3] := Binding_1_channels[2].retVal;
   TraceOut_channels_2_outputValue[3] := Binding_1_channels[2].outputValue;
   TraceOut_channels_3_enable[3] := Binding_1_channels[3].enable;
   TraceOut_channels_3_hiLIM[3] := Binding_1_channels[3].hiLIM;
   TraceOut_channels_3_loLIM[3] := Binding_1_channels[3].loLIM;
   TraceOut_channels_3_bipolar[3] := Binding_1_channels[3].bipolar;
   TraceOut_channels_3_measuringMode[3] := Binding_1_channels[3].measuringMode;
   TraceOut_channels_3_retVal[3] := Binding_1_channels[3].retVal;
   TraceOut_channels_3_outputValue[3] := Binding_1_channels[3].outputValue;
   TraceOut_channels_4_enable[3] := Binding_1_channels[4].enable;
   TraceOut_channels_4_hiLIM[3] := Binding_1_channels[4].hiLIM;
   TraceOut_channels_4_loLIM[3] := Binding_1_channels[4].loLIM;
   TraceOut_channels_4_bipolar[3] := Binding_1_channels[4].bipolar;
   TraceOut_channels_4_measuringMode[3] := Binding_1_channels[4].measuringMode;
   TraceOut_channels_4_retVal[3] := Binding_1_channels[4].retVal;
   TraceOut_channels_4_outputValue[3] := Binding_1_channels[4].outputValue;
   TraceOut_channels_5_enable[3] := Binding_1_channels[5].enable;
   TraceOut_channels_5_hiLIM[3] := Binding_1_channels[5].hiLIM;
   TraceOut_channels_5_loLIM[3] := Binding_1_channels[5].loLIM;
   TraceOut_channels_5_bipolar[3] := Binding_1_channels[5].bipolar;
   TraceOut_channels_5_measuringMode[3] := Binding_1_channels[5].measuringMode;
   TraceOut_channels_5_retVal[3] := Binding_1_channels[5].retVal;
   TraceOut_channels_5_outputValue[3] := Binding_1_channels[5].outputValue;
   TraceOut_channels_6_enable[3] := Binding_1_channels[6].enable;
   TraceOut_channels_6_hiLIM[3] := Binding_1_channels[6].hiLIM;
   TraceOut_channels_6_loLIM[3] := Binding_1_channels[6].loLIM;
   TraceOut_channels_6_bipolar[3] := Binding_1_channels[6].bipolar;
   TraceOut_channels_6_measuringMode[3] := Binding_1_channels[6].measuringMode;
   TraceOut_channels_6_retVal[3] := Binding_1_channels[6].retVal;
   TraceOut_channels_6_outputValue[3] := Binding_1_channels[6].outputValue;
   TraceOut_channels_7_enable[3] := Binding_1_channels[7].enable;
   TraceOut_channels_7_hiLIM[3] := Binding_1_channels[7].hiLIM;
   TraceOut_channels_7_loLIM[3] := Binding_1_channels[7].loLIM;
   TraceOut_channels_7_bipolar[3] := Binding_1_channels[7].bipolar;
   TraceOut_channels_7_measuringMode[3] := Binding_1_channels[7].measuringMode;
   TraceOut_channels_7_retVal[3] := Binding_1_channels[7].retVal;
   TraceOut_channels_7_outputValue[3] := Binding_1_channels[7].outputValue;
   TraceOut_channels_8_enable[3] := Binding_1_channels[8].enable;
   TraceOut_channels_8_hiLIM[3] := Binding_1_channels[8].hiLIM;
   TraceOut_channels_8_loLIM[3] := Binding_1_channels[8].loLIM;
   TraceOut_channels_8_bipolar[3] := Binding_1_channels[8].bipolar;
   TraceOut_channels_8_measuringMode[3] := Binding_1_channels[8].measuringMode;
   TraceOut_channels_8_retVal[3] := Binding_1_channels[8].retVal;
   TraceOut_channels_8_outputValue[3] := Binding_1_channels[8].outputValue;
   TraceOut_channels_9_enable[3] := Binding_1_channels[9].enable;
   TraceOut_channels_9_hiLIM[3] := Binding_1_channels[9].hiLIM;
   TraceOut_channels_9_loLIM[3] := Binding_1_channels[9].loLIM;
   TraceOut_channels_9_bipolar[3] := Binding_1_channels[9].bipolar;
   TraceOut_channels_9_measuringMode[3] := Binding_1_channels[9].measuringMode;
   TraceOut_channels_9_retVal[3] := Binding_1_channels[9].retVal;
   TraceOut_channels_9_outputValue[3] := Binding_1_channels[9].outputValue;
   BenchCalls := BenchCalls + 1;
 END_CASE;
 BenchStep := BenchStep + 1;
 IF BenchStep >= 4 THEN BenchDone := TRUE; END_IF;
END_IF;
END_PROGRAM
